// Device/Application/Equipment/FB_VacuumGripper
(*
    FB_VacuumGripper
    Purpose : Suction gripper: valve control with grip and loss supervision.
    Inputs  : xCmdVacuum, xVacuumOk (vacuum switch), tGripTimeout, itfAlarms
    Outputs : xValveOn, xHolding (vacuum on and OK)
    Errors  : VacuumNoGrip - commanded but not OK within tGripTimeout
              VacuumLost - was holding and lost vacuum while still commanded
*)
FUNCTION_BLOCK FB_VacuumGripper IMPLEMENTS I_Equipment
VAR_INPUT
    xCmdVacuum : BOOL;
    xVacuumOk : BOOL;
    tGripTimeout : TIME := T#500MS;
    itfAlarms : I_AlarmSink;
END_VAR
VAR_OUTPUT
    xValveOn : BOOL;
    xHolding : BOOL;
END_VAR
VAR
    tonGrip : TON;
    xWasHolding : BOOL;
    eError : E_AlarmId;
END_VAR

xValveOn := xCmdVacuum;
xHolding := xCmdVacuum AND xVacuumOk;

tonGrip(IN := xCmdVacuum AND NOT xVacuumOk AND NOT xWasHolding, PT := tGripTimeout);
IF tonGrip.Q AND eError = E_AlarmId.None THEN
    eError := E_AlarmId.VacuumNoGrip;
END_IF
IF xWasHolding AND xCmdVacuum AND NOT xVacuumOk AND eError = E_AlarmId.None THEN
    eError := E_AlarmId.VacuumLost;
END_IF

IF xHolding THEN
    xWasHolding := TRUE;
ELSIF NOT xCmdVacuum THEN
    xWasHolding := FALSE;
END_IF

IF eError <> E_AlarmId.None AND itfAlarms <> 0 THEN
    itfAlarms.Raise(eError);
END_IF

METHOD Reset : BOOL
IF itfAlarms <> 0 AND eError <> E_AlarmId.None THEN
    itfAlarms.Clear(eError);
END_IF
eError := E_AlarmId.None;
xWasHolding := FALSE;
Reset := TRUE;
END_METHOD

PROPERTY HasError : BOOL
GET
HasError := eError <> E_AlarmId.None;
END_GET
END_PROPERTY

PROPERTY ErrorId : E_AlarmId
GET
ErrorId := eError;
END_GET
END_PROPERTY

END_FUNCTION_BLOCK

// Device/Application/Equipment/FB_Bin
(*
    FB_Bin
    Purpose : Output bin: counts placed parts and reports the full sensor.
    Inputs  : eBin - which bin; xFullSensor; xPlaced - rising edge = one part placed
    Outputs : uiCount, xFull
    Methods : Empty() - operator emptied the bin
*)
FUNCTION_BLOCK FB_Bin
VAR_INPUT
    eBin : E_Bin;
    xFullSensor : BOOL;
    xPlaced : BOOL;
END_VAR
VAR_OUTPUT
    uiCount : UINT;
    xFull : BOOL;
END_VAR
VAR
    rtPlaced : R_TRIG;
END_VAR

rtPlaced(CLK := xPlaced);
IF rtPlaced.Q THEN
    uiCount := uiCount + 1;
END_IF
xFull := xFullSensor;

METHOD Empty
uiCount := 0;
END_METHOD

END_FUNCTION_BLOCK

// Device/Application/Equipment/FB_PhotoEye
(*
    FB_PhotoEye
    Purpose : Debounced photo-eye with a rising-edge pulse.
    Inputs  : xRaw - sensor signal (TRUE = beam blocked); tDebounce - on/off filter time
    Outputs : xBlocked - debounced state; xRising - TRUE for one cycle when it becomes blocked
*)
FUNCTION_BLOCK FB_PhotoEye
VAR_INPUT
    xRaw : BOOL;
    tDebounce : TIME := T#10MS;
END_VAR
VAR_OUTPUT
    xBlocked : BOOL;
    xRising : BOOL;
END_VAR
VAR
    tonOn : TON;
    tonOff : TON;
END_VAR

tonOn(IN := xRaw, PT := tDebounce);
tonOff(IN := NOT xRaw, PT := tDebounce);
xRising := FALSE;
IF tonOn.Q AND NOT xBlocked THEN
    xBlocked := TRUE;
    xRising := TRUE;
ELSIF tonOff.Q THEN
    xBlocked := FALSE;
END_IF

END_FUNCTION_BLOCK

// Device/Application/Comm/FB_BridgeWatchdog
(*
    FB_BridgeWatchdog
    Purpose : The Python bridge toggles xHeartbeat every cycle; if it stops toggling for tTimeout
              while enabled, the connection to the digital twin is considered lost.
    Outputs : xLost
    Alarms  : BridgeLost (Critical -> the cell aborts)
*)
FUNCTION_BLOCK FB_BridgeWatchdog
VAR_INPUT
    xHeartbeat : BOOL;
    xEnable : BOOL;
    tTimeout : TIME := T#500MS;
    itfAlarms : I_AlarmSink;
END_VAR
VAR_OUTPUT
    xLost : BOOL;
END_VAR
VAR
    xLastHeartbeat : BOOL;
    tonLost : TON;
END_VAR

tonLost(IN := xEnable AND xHeartbeat = xLastHeartbeat, PT := tTimeout);
xLastHeartbeat := xHeartbeat;
xLost := tonLost.Q;
IF itfAlarms <> 0 THEN
    IF xLost THEN
        itfAlarms.Raise(E_AlarmId.BridgeLost);
    ELSE
        itfAlarms.Clear(E_AlarmId.BridgeLost);
    END_IF
END_IF

END_FUNCTION_BLOCK

// Device/Application/Hmi/FB_HmiPanel
(*
    FB_HmiPanel
    Purpose : Turns the operator panel (GVL_HmiPanel: buttons, mode selector) into the cell's
              commands (GVL_Hmi). A button acts on its rising edge and is cleared, so a held or
              stuck button cannot repeat a command; the PackML state machine rejects commands
              that are not allowed in the current state.
    Inputs  : GVL_HmiPanel (written by the visualization), GVL_Bridge.eState
    Outputs : GVL_Hmi.eCommand / eModeRequest / xAlarmAck
    Modes   : iModeSelect 1 Production, 2 Maintenance, 3 Manual; other values are ignored. An
              operator change is requested only where PackML accepts a mode change (Stopped,
              Idle, Aborted), so no request waits to take effect after a later abort. The
              selector then shows GVL_Hmi.eModeRequest, whoever wrote it (panel or OPC UA).
*)
FUNCTION_BLOCK FB_HmiPanel
VAR
    rtStart : R_TRIG;
    rtStop : R_TRIG;
    rtReset : R_TRIG;
    rtClear : R_TRIG;
    rtAbort : R_TRIG;
    rtSuspend : R_TRIG;
    rtUnsuspend : R_TRIG;
    rtAck : R_TRIG;
    iLastMode : INT := 1;  // the selector value the panel showed last cycle
    xModeChangeAllowed : BOOL;
END_VAR

rtStart(CLK := GVL_HmiPanel.xStart);
rtStop(CLK := GVL_HmiPanel.xStop);
rtReset(CLK := GVL_HmiPanel.xReset);
rtClear(CLK := GVL_HmiPanel.xClear);
rtAbort(CLK := GVL_HmiPanel.xAbort);
rtSuspend(CLK := GVL_HmiPanel.xSuspend);
rtUnsuspend(CLK := GVL_HmiPanel.xUnsuspend);
rtAck(CLK := GVL_HmiPanel.xAckAll);

// Abort and Stop first: a safety-relevant command wins over a start in the same cycle.
IF rtAbort.Q THEN
    GVL_Hmi.eCommand := E_PackMLCommand.Abort;
ELSIF rtStop.Q THEN
    GVL_Hmi.eCommand := E_PackMLCommand.Stop;
ELSIF rtClear.Q THEN
    GVL_Hmi.eCommand := E_PackMLCommand.Clear;
ELSIF rtReset.Q THEN
    GVL_Hmi.eCommand := E_PackMLCommand.Reset;
ELSIF rtSuspend.Q THEN
    GVL_Hmi.eCommand := E_PackMLCommand.Suspend;
ELSIF rtUnsuspend.Q THEN
    GVL_Hmi.eCommand := E_PackMLCommand.Unsuspend;
ELSIF rtStart.Q THEN
    GVL_Hmi.eCommand := E_PackMLCommand.Start;
END_IF
IF rtAck.Q THEN
    GVL_Hmi.xAlarmAck := TRUE;
END_IF

// mode selector: an operator change, only where PackML accepts it
IF GVL_HmiPanel.iModeSelect <> iLastMode THEN
    xModeChangeAllowed := GVL_Bridge.eState = E_PackMLState.Stopped
                          OR GVL_Bridge.eState = E_PackMLState.Idle
                          OR GVL_Bridge.eState = E_PackMLState.Aborted;
    IF xModeChangeAllowed THEN
        CASE GVL_HmiPanel.iModeSelect OF
            1: GVL_Hmi.eModeRequest := E_PackMLMode.Production;
            2: GVL_Hmi.eModeRequest := E_PackMLMode.Maintenance;
            3: GVL_Hmi.eModeRequest := E_PackMLMode.Manual;
        END_CASE   // other values: ignored
    END_IF
END_IF
// the selector shows the request (refused or invalid choices fall back, OPC UA requests show)
CASE GVL_Hmi.eModeRequest OF
    E_PackMLMode.Production: iLastMode := 1;
    E_PackMLMode.Maintenance: iLastMode := 2;
    E_PackMLMode.Manual: iLastMode := 3;
END_CASE
GVL_HmiPanel.iModeSelect := iLastMode;

GVL_HmiPanel.xStart := FALSE;
GVL_HmiPanel.xStop := FALSE;
GVL_HmiPanel.xReset := FALSE;
GVL_HmiPanel.xClear := FALSE;
GVL_HmiPanel.xAbort := FALSE;
GVL_HmiPanel.xSuspend := FALSE;
GVL_HmiPanel.xUnsuspend := FALSE;
GVL_HmiPanel.xAckAll := FALSE;

END_FUNCTION_BLOCK

// Device/Application/Hmi/FB_HmiView
(*
    FB_HmiView
    Purpose : Prepares the display data of the visualization (GVL_HmiView): state and mode texts,
              state groups for the machine bar, alarm rows (active or unacknowledged, and the
              condition itself), newest alarm text, equipment signals and the placed counter.
    In/Out  : Cell - the sorting cell (read only)
    Outputs : GVL_HmiView
*)
FUNCTION_BLOCK FB_HmiView
VAR_IN_OUT
    Cell : FB_SortingCell;
END_VAR
VAR
    i : INT;
    stAlarm : ST_Alarm;
END_VAR
VAR CONSTANT
    BELT_RUNNING_MM_S : LREAL := 1.0;  // the belt counts as running above this speed
    // HMI row i shows alarm ALARM_ROWS[i] (E_AlarmId is strict: no integer arithmetic on it)
    ALARM_ROWS : ARRAY[1..16] OF E_AlarmId := [
        E_AlarmId.EStop, E_AlarmId.DoorOpen, E_AlarmId.BridgeLost, E_AlarmId.AxisGroupError,
        E_AlarmId.ConveyorError, E_AlarmId.FollowingErrorWarn, E_AlarmId.FollowingErrorFault,
        E_AlarmId.FeedbackStale, E_AlarmId.VacuumNoGrip, E_AlarmId.VacuumLost,
        E_AlarmId.PartMissed, E_AlarmId.BinFull, E_AlarmId.VisionMissing,
        E_AlarmId.DecisionFallback, E_AlarmId.LowConfidence, E_AlarmId.QueueOverflow];
END_VAR

CASE Cell.eState OF
    E_PackMLState.Clearing: GVL_HmiView.sState := 'Clearing';
    E_PackMLState.Stopped: GVL_HmiView.sState := 'Stopped';
    E_PackMLState.Starting: GVL_HmiView.sState := 'Starting';
    E_PackMLState.Idle: GVL_HmiView.sState := 'Idle';
    E_PackMLState.Suspended: GVL_HmiView.sState := 'Suspended';
    E_PackMLState.Execute: GVL_HmiView.sState := 'Execute';
    E_PackMLState.Stopping: GVL_HmiView.sState := 'Stopping';
    E_PackMLState.Aborting: GVL_HmiView.sState := 'Aborting';
    E_PackMLState.Aborted: GVL_HmiView.sState := 'Aborted';
    E_PackMLState.Holding: GVL_HmiView.sState := 'Holding';
    E_PackMLState.Held: GVL_HmiView.sState := 'Held';
    E_PackMLState.Unholding: GVL_HmiView.sState := 'Unholding';
    E_PackMLState.Suspending: GVL_HmiView.sState := 'Suspending';
    E_PackMLState.Unsuspending: GVL_HmiView.sState := 'Unsuspending';
    E_PackMLState.Resetting: GVL_HmiView.sState := 'Resetting';
    E_PackMLState.Completing: GVL_HmiView.sState := 'Completing';
    E_PackMLState.Complete: GVL_HmiView.sState := 'Complete';
ELSE
    GVL_HmiView.sState := 'Undefined';
END_CASE
CASE Cell.eMode OF
    E_PackMLMode.Production: GVL_HmiView.sMode := 'Production';
    E_PackMLMode.Maintenance: GVL_HmiView.sMode := 'Maintenance';
    E_PackMLMode.Manual: GVL_HmiView.sMode := 'Manual';
END_CASE
CASE Cell.ePickStep OF
    E_PickStep.Idle: GVL_HmiView.sPickStep := 'Idle';
    E_PickStep.MoveHome: GVL_HmiView.sPickStep := 'Moving home';
    E_PickStep.MoveReady: GVL_HmiView.sPickStep := 'Moving to ready';
    E_PickStep.WaitPart: GVL_HmiView.sPickStep := 'Waiting for a part';
    E_PickStep.StartTracking: GVL_HmiView.sPickStep := 'Tracking the belt';
    E_PickStep.Approach: GVL_HmiView.sPickStep := 'Approaching';
    E_PickStep.Descend: GVL_HmiView.sPickStep := 'Descending';
    E_PickStep.Grip: GVL_HmiView.sPickStep := 'Gripping';
    E_PickStep.Lift: GVL_HmiView.sPickStep := 'Lifting';
    E_PickStep.MoveToBin: GVL_HmiView.sPickStep := 'Moving to bin';
    E_PickStep.Release: GVL_HmiView.sPickStep := 'Releasing';
    E_PickStep.Retract: GVL_HmiView.sPickStep := 'Retracting';
    E_PickStep.Aborting: GVL_HmiView.sPickStep := 'Stopping';
    E_PickStep.Aborted: GVL_HmiView.sPickStep := 'Stopped (abort)';
    E_PickStep.Error: GVL_HmiView.sPickStep := 'Error';
    E_PickStep.RecoverLift: GVL_HmiView.sPickStep := 'Recovering';
END_CASE

GVL_HmiView.xExecute := Cell.eState = E_PackMLState.Execute;
GVL_HmiView.xStopped := Cell.eState = E_PackMLState.Stopped;
GVL_HmiView.xIdle := Cell.eState = E_PackMLState.Idle;
GVL_HmiView.xAborted := Cell.eState = E_PackMLState.Aborted OR Cell.eState = E_PackMLState.Aborting;
GVL_HmiView.xHeld := Cell.eState = E_PackMLState.Held OR Cell.eState = E_PackMLState.Suspended
                     OR Cell.eState = E_PackMLState.Holding OR Cell.eState = E_PackMLState.Suspending;
GVL_HmiView.xActing := Cell.eState = E_PackMLState.Resetting OR Cell.eState = E_PackMLState.Starting
                       OR Cell.eState = E_PackMLState.Stopping OR Cell.eState = E_PackMLState.Clearing
                       OR Cell.eState = E_PackMLState.Unholding OR Cell.eState = E_PackMLState.Unsuspending;
GVL_HmiView.xManual := Cell.eMode = E_PackMLMode.Manual;
GVL_HmiView.xJogPermitted := GVL_HmiView.xManual AND GVL_HmiView.xExecute;

GVL_HmiView.xAnyAlarm := FALSE;
FOR i := 1 TO 16 DO
    stAlarm := Cell.AlarmState(ALARM_ROWS[i]);
    GVL_HmiView.axAlarmActive[i] := stAlarm.xActive;
    GVL_HmiView.axAlarm[i] := stAlarm.xActive OR NOT stAlarm.xAcked;
    GVL_HmiView.xAnyAlarm := GVL_HmiView.xAnyAlarm OR GVL_HmiView.axAlarm[i];
END_FOR
GVL_HmiView.sNewestAlarm := GVL_AlarmDefs.aDefs[Cell.eNewestAlarm].sText;
GVL_HmiView.uiPlaced := Cell.PlacedCount();
GVL_HmiView.xBeltRunning := ABS(Cell.lrBeltVel) > BELT_RUNNING_MM_S;
GVL_HmiView.xRobotMoving := Cell.RobotMoving();
GVL_HmiView.xAnyBinFull := Cell.AnyBinFull();

END_FUNCTION_BLOCK

// Device/Application/Tests/PRG_Tests
(*
    PRG_Tests
    Purpose : Calls every simulation test harness (TEST programs in this folder).
    Task    : TestTask, cyclic 10 ms
*)
PROGRAM PRG_Tests
VAR
END_VAR

PRG_TestMotionSmoke();
PRG_TestTypes();
PRG_TestPackML();
PRG_TestAlarms();
PRG_TestEquipment();
PRG_TestMotion();
PRG_TestJointMonitor();
PRG_TestTracking();
PRG_TestPick();
PRG_TestCell();

END_PROGRAM

// Device/Application/Tests/PRG_TestMotionSmoke
(*
    PRG_TestMotionSmoke
    Purpose : Simulation test harness - powers the robot axis group and makes one PTP move.
    Task    : TestTask (via PRG_Tests)
    Spec    : tests/plc/motion_smoke.json
*)
PROGRAM PRG_TestMotionSmoke
VAR
    fbPower : SMC_GroupPower;
    fbEnable : MC_GroupEnable;
    fbMove : MC_MoveDirectAbsolute := (CoordSystem := SMC_COORD_SYSTEM.ACS, VelFactor := 0.5);
    fbReadPos : MC_GroupReadActualPosition := (Enable := TRUE, CoordSystem := SMC_COORD_SYSTEM.ACS);
    xGo : BOOL;
    lrJ1 : LREAL;
    lrJ2 : LREAL;
    xMoveDone : BOOL;
    xMoveError : BOOL;
END_VAR

// Only commands the robot while the test runs, so other harnesses can use it.
IF xGo THEN
    fbPower(AxisGroup := AxisGroup_Robot, Enable := TRUE, bRegulatorOn := TRUE, bDriveStart := TRUE);
    fbEnable(AxisGroup := AxisGroup_Robot, Execute := fbPower.Status);
    fbMove.Position.a.a0 := 30;
    fbMove.Position.a.a1 := -20;
    fbMove.Position.a.a2 := 40;
    fbMove.Position.a.a3 := 0;
    fbMove.Position.a.a4 := 45;
    fbMove.Position.a.a5 := 0;
    fbMove(AxisGroup := AxisGroup_Robot, Execute := fbEnable.Done);
    fbReadPos(AxisGroup := AxisGroup_Robot);
    lrJ1 := fbReadPos.Position.a.a0;
    lrJ2 := fbReadPos.Position.a.a1;
    xMoveDone := fbMove.Done;
    xMoveError := fbMove.Error;
END_IF

END_PROGRAM

// Device/Application/Tests/PRG_TestTypes
(*
    PRG_TestTypes
    Purpose : Simulation test harness - exposes configuration values for tests/plc/types.json.
*)
PROGRAM PRG_TestTypes
VAR
    eClassBin0 : E_Bin;
    eFaultClass : E_AlarmClass;
    eWarnClass : E_AlarmClass;
    xLoopback : BOOL;
END_VAR

eClassBin0 := GVL_Params.aClassToBin[0];
eFaultClass := GVL_AlarmDefs.aDefs[E_AlarmId.EStop].eClass;
eWarnClass := GVL_AlarmDefs.aDefs[E_AlarmId.PartMissed].eClass;
xLoopback := GVL_Config.xFeedbackLoopback;

END_PROGRAM

// Device/Application/Tests/PRG_TestPackML
(*
    PRG_TestPackML
    Purpose : Simulation test harness for FB_PackMLStateMachine (tests/plc/packml.json).
    Inputs  : xReinit - TRUE re-initialises the state machine, then resets itself.
*)
PROGRAM PRG_TestPackML
VAR
    fbSm : FB_PackMLStateMachine;
    fbSmInitial : FB_PackMLStateMachine;
    xReinit : BOOL;
END_VAR

IF xReinit THEN
    xReinit := FALSE;
    fbSm := fbSmInitial;
END_IF
fbSm();

END_PROGRAM

// Device/Application/Tests/PRG_TestAlarms
(*
    PRG_TestAlarms
    Purpose : Simulation test harness for FB_AlarmHandler (tests/plc/alarms.json).
    Inputs  : eId + xRaise / xRaiseEvent / xClear pulses, xAck, xReinit (each pulse resets itself).
*)
PROGRAM PRG_TestAlarms
VAR
    fbAlarms : FB_AlarmHandler;
    fbAlarmsInitial : FB_AlarmHandler;
    eId : E_AlarmId;
    xRaise : BOOL;
    xRaiseEvent : BOOL;
    xClear : BOOL;
    xAck : BOOL;
    xReinit : BOOL;
END_VAR

IF xReinit THEN
    xReinit := FALSE;
    fbAlarms := fbAlarmsInitial;
END_IF
IF xRaise THEN
    xRaise := FALSE;
    fbAlarms.Raise(eId);
END_IF
IF xRaiseEvent THEN
    xRaiseEvent := FALSE;
    fbAlarms.RaiseEvent(eId);
END_IF
IF xClear THEN
    xClear := FALSE;
    fbAlarms.Clear(eId);
END_IF
IF xAck THEN
    xAck := FALSE;
    fbAlarms.AcknowledgeAll();
END_IF
fbAlarms();

END_PROGRAM

// Device/Application/Tests/PRG_TestEquipment
(*
    PRG_TestEquipment
    Purpose : Simulation test harness for the simple equipment FBs (tests/plc/equipment.json).
    Pulses  : write udiPulseMs and set xStartPulse - the harness drives fbPe.xRaw for exactly
              that long in PLC time (tool writes are too slow to time a short pulse).
*)
PROGRAM PRG_TestEquipment
VAR
    fbAlarms : FB_AlarmHandler;
    fbPe : FB_PhotoEye := (tDebounce := T#300MS);
    fbVac : FB_VacuumGripper;
    fbBin : FB_Bin := (eBin := E_Bin.TypeA);
    fbSafety : FB_SafetyMonitor;
    fbAlarmsInitial : FB_AlarmHandler;
    fbPeInitial : FB_PhotoEye := (tDebounce := T#300MS);
    fbVacInitial : FB_VacuumGripper;
    fbBinInitial : FB_Bin := (eBin := E_Bin.TypeA);
    fbSafetyInitial : FB_SafetyMonitor;
    xReinit : BOOL;
    uiPeRises : UINT;
    eVacError : E_AlarmId;
    udiPulseMs : UDINT;
    xStartPulse : BOOL;
    xPulseActive : BOOL;
    tonPulse : TON;
END_VAR

IF xReinit THEN
    xReinit := FALSE;
    fbAlarms := fbAlarmsInitial;
    fbPe := fbPeInitial;
    fbVac := fbVacInitial;
    fbBin := fbBinInitial;
    fbSafety := fbSafetyInitial;
    uiPeRises := 0;
    xPulseActive := FALSE;
END_IF
fbVac.itfAlarms := fbAlarms;
fbSafety.itfAlarms := fbAlarms;

IF xStartPulse THEN
    xStartPulse := FALSE;
    xPulseActive := TRUE;
END_IF
tonPulse(IN := xPulseActive, PT := TO_TIME(udiPulseMs));
IF tonPulse.Q THEN
    xPulseActive := FALSE;
END_IF
fbPe.xRaw := xPulseActive;

fbPe();
IF fbPe.xRising THEN
    uiPeRises := uiPeRises + 1;
END_IF
fbVac();
eVacError := fbVac.ErrorId;
fbBin();
fbSafety();
fbAlarms();

END_PROGRAM

// Device/Application/Tests/PRG_TestMotion
(*
    PRG_TestMotion
    Purpose : Simulation test harness for FB_Robot and FB_Conveyor (tests/plc/motion.json).
    Inputs  : xActive - only then are the FBs called; xGo - start eCmd with the target chosen by
              iTargetSel (1 = home, 2 = current TCP - 50 mm in Z, 3 = home with J1 = 60 deg,
              4 = stProbe as written by the test)
    Outputs : xLastDone / xLastError of the last command, udiMoveMsLast / udiMoveMsPrev,
              xSlower (last move took > 1.5 x the previous one), lrZDelta
    Note    : SoftMotion FB instances are never re-initialised by assignment (corrupts them).
*)
PROGRAM PRG_TestMotion
VAR
    fbRobot : FB_Robot;
    fbConv : FB_Conveyor;
    fbAlarms : FB_AlarmHandler;
    xActive : BOOL;
    iTargetSel : INT;
    eCmd : E_RobotCmd;
    xGo : BOOL;
    iGoStep : INT;
    xLastDone : BOOL;
    xLastError : BOOL;
    tStart : TIME;
    udiMoveMsLast : UDINT;
    udiMoveMsPrev : UDINT;
    xSlower : BOOL;
    lrZStart : LREAL;
    lrZDelta : LREAL;
    stTarget : SMC_POS_REF;
    stProbe : SMC_POS_REF;
END_VAR

IF NOT xActive THEN
    RETURN;
END_IF
fbRobot.itfAlarms := fbAlarms;
fbConv.itfAlarms := fbAlarms;

IF xGo THEN
    xGo := FALSE;
    CASE iTargetSel OF
        1: stTarget := GVL_CellGeometry.HOME_ACS;
        2: stTarget := fbRobot.stActMcs;
           lrZStart := fbRobot.stActMcs.c.Z;
           stTarget.c.Z := lrZStart - 50;
        3: stTarget := GVL_CellGeometry.HOME_ACS;
           stTarget.a.a0 := 60;
        4: stTarget := stProbe;
    END_CASE
    fbRobot.stTarget := stTarget;
    fbRobot.eCmd := eCmd;
    fbRobot.xExecute := FALSE;     // a fresh rising edge, even if a command is running
    iGoStep := 1;
    xLastDone := FALSE;
    xLastError := FALSE;
ELSIF iGoStep = 1 THEN
    fbRobot.xExecute := TRUE;
    tStart := TIME();
    iGoStep := 2;
ELSIF iGoStep = 2 AND (fbRobot.xDone OR fbRobot.xError) THEN
    xLastDone := fbRobot.xDone;
    xLastError := fbRobot.xError;
    udiMoveMsPrev := udiMoveMsLast;
    udiMoveMsLast := TIME_TO_UDINT(TIME() - tStart);
    xSlower := udiMoveMsLast * 2 > udiMoveMsPrev * 3;
    fbRobot.xExecute := FALSE;
    iGoStep := 0;
END_IF

fbRobot(AxisGroup := AxisGroup_Robot);
fbConv(Axis := Axis_Conveyor);
fbAlarms();
IF iTargetSel = 2 THEN
    lrZDelta := fbRobot.stActMcs.c.Z - lrZStart;
END_IF

END_PROGRAM

// Device/Application/Tests/PRG_TestJointMonitor
(*
    PRG_TestJointMonitor
    Purpose : Simulation test harness for FB_JointMonitor (tests/plc/joint_monitor.json).
    Inputs  : xReinit; xAutoSeq - increment the feedback and setpoint sequences every cycle
              xRamp - J1 setpoint ramps by RAMP_STEP per cycle; iLag - feedback is the setpoint of
              iLag cycles earlier (and says so in udiFeedbackForSeq); xFreeze - feedback stands still;
              iTornSamples - that many cycles claim a sample iTornAge older (a torn OPC UA write,
              or a bridge hiccup when iTornAge exceeds the history)
    Outputs : lrRampSpeed - measured J1 setpoint speed [deg/s]
*)
PROGRAM PRG_TestJointMonitor
VAR
    fbMon : FB_JointMonitor;
    fbAlarms : FB_AlarmHandler;
    fbMonInitial : FB_JointMonitor;
    fbAlarmsInitial : FB_AlarmHandler;
    xReinit : BOOL;
    xAutoSeq : BOOL;
    xRamp : BOOL;
    xFreeze : BOOL;
    iLag : INT;
    udiSpSeq : UDINT;
    aSpHist : ARRAY[0..127] OF LREAL;
    xRampOld : BOOL;
    tRampStart : TIME;
    lrRampStart : LREAL;
    lrRampSpeed : LREAL;
    iTornSamples : INT;             // next cycles: feedback says it answers an older sample
    iTornAge : INT := 25;           // [samples]
END_VAR
VAR CONSTANT
    RAMP_STEP : LREAL := 1.0;       // [deg per cycle]
END_VAR

IF xReinit THEN
    xReinit := FALSE;
    xAutoSeq := FALSE;
    xRamp := FALSE;
    xFreeze := FALSE;
    iLag := 0;
    iTornSamples := 0;
    udiSpSeq := 0;
    fbMon := fbMonInitial;
    fbAlarms := fbAlarmsInitial;
END_IF
IF xAutoSeq THEN
    fbMon.udiFeedbackSeq := fbMon.udiFeedbackSeq + 1;
    udiSpSeq := udiSpSeq + 1;
END_IF
IF xRamp THEN
    IF NOT xRampOld THEN
        tRampStart := TIME();
        lrRampStart := fbMon.aSetpoint[1];
    END_IF
    fbMon.aSetpoint[1] := fbMon.aSetpoint[1] + RAMP_STEP;
    IF TIME() > tRampStart THEN
        lrRampSpeed := (fbMon.aSetpoint[1] - lrRampStart) * 1000.0 / TIME_TO_LREAL(TIME() - tRampStart);
    END_IF
END_IF
xRampOld := xRamp;
aSpHist[udiSpSeq MOD 128] := fbMon.aSetpoint[1];
fbMon.udiSetpointSeq := udiSpSeq;
IF udiSpSeq >= INT_TO_UDINT(iLag) THEN
    fbMon.udiFeedbackForSeq := udiSpSeq - INT_TO_UDINT(iLag);
    IF NOT xFreeze THEN
        fbMon.aFeedback[1] := aSpHist[fbMon.udiFeedbackForSeq MOD 128];
    END_IF
    IF iTornSamples > 0 AND fbMon.udiFeedbackForSeq >= INT_TO_UDINT(iTornAge) THEN
        fbMon.udiFeedbackForSeq := fbMon.udiFeedbackForSeq - INT_TO_UDINT(iTornAge);
        iTornSamples := iTornSamples - 1;
    END_IF
END_IF
fbMon.itfAlarms := fbAlarms;
fbMon();
fbAlarms();

END_PROGRAM

// Device/Application/Tests/PRG_TestTracking
(*
    PRG_TestTracking
    Purpose : Simulation test harness for FB_PartTracker and F_SelectBin (tests/plc/tracking.json).
    Inputs  : lrBeltPos; xTriggerPE1 (one capture); uiFillCount (that many captures, one per cycle);
              stVisIn + xSendVision / xResendVision (same sequence number again);
              stDecIn + xSendDecision; udiQueryId - part to show in stRec; xAck; xClear;
              xNoDecisionLayer (no AI decision service)
    Outputs : uiCount, uiNext (next pickable index), stRec, xQueryFound
*)
PROGRAM PRG_TestTracking
VAR
    fbTracker : FB_PartTracker;
    fbAlarms : FB_AlarmHandler;
    fbTrackerInitial : FB_PartTracker;
    fbAlarmsInitial : FB_AlarmHandler;
    xReinit : BOOL;
    lrBeltPos : LREAL;
    xTriggerPE1 : BOOL;
    uiFillCount : UINT;
    stVisIn : ST_VisionMsg;
    stDecIn : ST_DecisionMsg;
    xSendVision : BOOL;
    xResendVision : BOOL;
    xSendDecision : BOOL;
    xAck : BOOL;
    xClear : BOOL;
    udiVisionSeq : UDINT;
    udiDecisionSeq : UDINT;
    udiQueryId : UDINT;
    uiQueryIdx : UINT;
    xQueryFound : BOOL;
    stRec : ST_PartRecord;
    uiCount : UINT;
    uiNext : UINT;
    xPE1Rising : BOOL;
    xNoDecisionLayer : BOOL;
END_VAR

IF xReinit THEN
    xReinit := FALSE;
    fbTracker := fbTrackerInitial;
    fbAlarms := fbAlarmsInitial;
    udiVisionSeq := 0;
    udiDecisionSeq := 0;
    uiFillCount := 0;
END_IF

xPE1Rising := xTriggerPE1 OR uiFillCount > 0;
xTriggerPE1 := FALSE;
IF uiFillCount > 0 THEN
    uiFillCount := uiFillCount - 1;
END_IF

IF xSendVision THEN
    xSendVision := FALSE;
    udiVisionSeq := udiVisionSeq + 1;
END_IF
IF xResendVision THEN
    xResendVision := FALSE;      // same sequence number: must be ignored
END_IF
stVisIn.udiSeq := udiVisionSeq;
IF xSendDecision THEN
    xSendDecision := FALSE;
    udiDecisionSeq := udiDecisionSeq + 1;
END_IF
stDecIn.udiSeq := udiDecisionSeq;
IF xAck THEN
    xAck := FALSE;
    fbAlarms.AcknowledgeAll();
END_IF
IF xClear THEN
    xClear := FALSE;
    fbTracker.Clear();
END_IF

fbTracker.itfAlarms := fbAlarms;
fbTracker(lrBeltPos := lrBeltPos, xPE1Rising := xPE1Rising, stVision := stVisIn, stDecision := stDecIn,
          xDecisionActive := NOT xNoDecisionLayer);
fbAlarms();

uiCount := fbTracker.Count;
uiNext := fbTracker.NextPickable(GVL_CellGeometry.PE2_X, GVL_CellGeometry.PICK_WINDOW_END_X);
uiQueryIdx := fbTracker.FindPart(udiQueryId);
xQueryFound := uiQueryIdx > 0;
IF xQueryFound THEN
    stRec := fbTracker.GetRecord(uiQueryIdx);
END_IF

END_PROGRAM

// Device/Application/Tests/PRG_TestPick
(*
    PRG_TestPick
    Purpose : Simulation test harness for FB_PickSequence (tests/plc/pick.json). Owns the robot,
              conveyor, gripper, tracker and alarms like the cell does, and simulates the vacuum
              switch (OK 100 ms after the valve opens).
    Inputs  : xActive, xBeltRun, xInject (+ usiInjClass, eInjQuality, lrInjX: one part with
              vision and decision; xInjInvalid: the vision message says "not seen"),
              xDropOnTransfer (vacuum lost during MoveToBin),
              xAbortOnLift (abort when the sequence reaches Lift), xResetSeq
    Outputs : xSawRecoverLift (latched: the recovery after an abort lifted first),
              lrGripZ (TCP height when the last grip started) [mm]
    Note    : SoftMotion FB instances are never re-initialised by assignment.
*)
PROGRAM PRG_TestPick
VAR
    fbRobot : FB_Robot;
    fbConv : FB_Conveyor;
    fbVac : FB_VacuumGripper;
    fbTracker : FB_PartTracker;
    fbAlarms : FB_AlarmHandler;
    fbSeq : FB_PickSequence;
    xActive : BOOL;
    xBeltRun : BOOL;
    xInject : BOOL;
    xInjInvalid : BOOL;
    usiInjClass : USINT;
    eInjQuality : E_Quality := E_Quality.Ok;
    lrInjX : LREAL := 1000;
    iInject : INT;
    xPE1 : BOOL;
    stVis : ST_VisionMsg;
    stDec : ST_DecisionMsg;
    xDropOnTransfer : BOOL;
    xAbortOnLift : BOOL;
    xResetSeq : BOOL;
    xVacLost : BOOL;
    tonVac : TON;
    xSawRecoverLift : BOOL;
    lrGripZ : LREAL;
    eLastStep : E_PickStep;
END_VAR

IF NOT xActive THEN
    RETURN;
END_IF
fbRobot.itfAlarms := fbAlarms;
fbConv.itfAlarms := fbAlarms;
fbVac.itfAlarms := fbAlarms;
fbTracker.itfAlarms := fbAlarms;
fbConv.xEnable := TRUE;
fbConv.lrVelocity := GVL_Params.lrBeltSpeed;
fbConv.xRun := xBeltRun;
fbRobot.xEnable := TRUE;

// One injected part: capture, then vision, then decision on consecutive cycles.
CASE iInject OF
    0:
        IF xInject THEN
            xInject := FALSE;
            xPE1 := TRUE;
            iInject := 1;
        END_IF
    1:
        xPE1 := FALSE;
        iInject := 2;
    2:
        stVis.udiSeq := stVis.udiSeq + 1;
        stVis.udiPartId := fbTracker.stCapture.udiPartId;
        stVis.xValid := NOT xInjInvalid;
        stVis.usiClass := usiInjClass;
        stVis.rConfidence := 0.9;
        stVis.lrX := lrInjX;
        stVis.lrY := 0;
        stVis.lrTheta := 0;
        iInject := 3;
    3:
        stDec.udiSeq := stDec.udiSeq + 1;
        stDec.udiPartId := stVis.udiPartId;
        stDec.eQuality := eInjQuality;
        stDec.rQualityProb := 0.95;
        stDec.xIdentReliable := TRUE;
        iInject := 0;
END_CASE

IF xDropOnTransfer AND fbSeq.eStep = E_PickStep.MoveToBin THEN
    xVacLost := TRUE;
END_IF
tonVac(IN := fbVac.xValveOn AND NOT xVacLost, PT := T#100MS);
fbVac.xVacuumOk := tonVac.Q;
IF xAbortOnLift AND fbSeq.eStep = E_PickStep.Lift THEN
    fbSeq.xAbort := TRUE;
END_IF
fbSeq.xReset := xResetSeq;
IF xResetSeq THEN
    xResetSeq := FALSE;
    xVacLost := FALSE;
    fbSeq.xAbort := FALSE;
    fbVac.Reset();
    fbAlarms.AcknowledgeAll();
END_IF

fbTracker(lrBeltPos := fbConv.lrPosition, xPE1Rising := xPE1, stVision := stVis, stDecision := stDec);
fbSeq(AxisGroup := AxisGroup_Robot, ConveyorAxis := Axis_Conveyor, Robot := fbRobot, Gripper := fbVac, Tracker := fbTracker);
fbVac();
fbRobot(AxisGroup := AxisGroup_Robot);
fbConv(Axis := Axis_Conveyor);
fbAlarms();
IF fbSeq.eStep = E_PickStep.RecoverLift THEN
    xSawRecoverLift := TRUE;
END_IF
IF fbSeq.eStep = E_PickStep.Grip AND eLastStep <> E_PickStep.Grip THEN
    lrGripZ := fbRobot.stActMcs.c.Z;
END_IF
eLastStep := fbSeq.eStep;

END_PROGRAM

// Device/Application/Tests/PRG_TestCell
(*
    PRG_TestCell
    Purpose : Simulation test harness for the whole cell in PRG_Main (tests/plc/cell.json).
              Simulates the vacuum switch, injects parts (PE1 pulse, then vision and decision
              messages for the captured part id) and can press the E-stop or lose the vacuum
              during a transfer. Can play the twin's bridge (heartbeat, joint feedback answering
              the current setpoint sample, twin active) and stall it. While active it plays an AI
              decision service (GVL_Bridge.xDecisionActive), reset when it is switched off.
    Inputs  : xActive; xInject (+ usiInjClass, eInjQuality); xEStopOnTransfer; xVacLostOnTransfer;
              xMark (J1 reference); xBridgeSim; xBridgeStall (heartbeat stops toggling);
              xBridgeStallOnTransfer
    Outputs : lrJ1Delta - J1 movement since xMark [deg]; lrAbortDelayMs - bridge stall -> Aborted
*)
PROGRAM PRG_TestCell
VAR
    xActive : BOOL;
    xWasActive : BOOL;
    xInject : BOOL;
    usiInjClass : USINT;
    eInjQuality : E_Quality := E_Quality.Ok;
    iInject : INT;
    tonPulse : TON;
    tonVac : TON;
    xEStopOnTransfer : BOOL;
    xVacLostOnTransfer : BOOL;
    xVacLost : BOOL;                    // latched until xVacLostOnTransfer is released
    xMark : BOOL;
    lrJ1Start : LREAL;
    lrJ1Delta : LREAL;
    xBridgeSim : BOOL;
    xBridgeStall : BOOL;
    xBridgeStallOnTransfer : BOOL;      // stall the bridge when the robot carries a part to its bin
    xStallTimed : BOOL;
    tStall : TIME;
    lrAbortDelayMs : LREAL;             // stall -> Aborted [ms]
END_VAR
VAR CONSTANT
    PE1_PULSE : TIME := T#250MS;
END_VAR

IF NOT xActive THEN
    IF xWasActive THEN                   // leave no fake decision service behind
        GVL_Bridge.xDecisionActive := FALSE;
        xWasActive := FALSE;
    END_IF
    RETURN;
END_IF
xWasActive := TRUE;
GVL_Bridge.xDecisionActive := TRUE;  // the harness injects AI decisions (eInjQuality)

IF xVacLostOnTransfer AND PRG_Main.fbCell.ePickStep = E_PickStep.MoveToBin THEN
    xVacLost := TRUE;
ELSIF NOT xVacLostOnTransfer THEN
    xVacLost := FALSE;
END_IF
tonVac(IN := GVL_Bridge.xVacuumOn, PT := T#100MS);
GVL_Bridge.xVacuumOk := tonVac.Q AND NOT xVacLost;

// the twin's bridge: feedback answers the current setpoint sample, heartbeat toggles
IF xBridgeStallOnTransfer AND NOT xBridgeStall AND PRG_Main.fbCell.ePickStep = E_PickStep.MoveToBin THEN
    xBridgeStall := TRUE;
    xStallTimed := FALSE;
    tStall := TIME();
END_IF
IF xBridgeStall AND NOT xStallTimed AND GVL_Bridge.eState = E_PackMLState.Aborted THEN
    xStallTimed := TRUE;
    lrAbortDelayMs := TIME_TO_LREAL(TIME() - tStall);
END_IF
IF xBridgeSim THEN
    GVL_Bridge.xTwinActive := TRUE;
    GVL_Bridge.aJointPosFb := GVL_Bridge.aJointPosSp;
    GVL_Bridge.udiFeedbackForSeq := GVL_Bridge.udiSetpointSeq;
    IF NOT xBridgeStall THEN
        GVL_Bridge.xHeartbeat := NOT GVL_Bridge.xHeartbeat;
        GVL_Bridge.udiFeedbackSeq := GVL_Bridge.udiFeedbackSeq + 1;
    END_IF
END_IF

CASE iInject OF
    0:
        IF xInject THEN
            xInject := FALSE;
            GVL_Bridge.xPE1 := TRUE;
            iInject := 1;
        END_IF
    1:
        tonPulse(IN := TRUE, PT := PE1_PULSE);
        IF tonPulse.Q THEN
            tonPulse(IN := FALSE);
            GVL_Bridge.xPE1 := FALSE;
            iInject := 2;
        END_IF
    2:
        GVL_Bridge.stVision.udiPartId := GVL_Bridge.stCapture.udiPartId;
        GVL_Bridge.stVision.xValid := TRUE;
        GVL_Bridge.stVision.usiClass := usiInjClass;
        GVL_Bridge.stVision.rConfidence := 0.9;
        GVL_Bridge.stVision.lrX := GVL_CellGeometry.PE1_X;
        GVL_Bridge.stVision.lrY := 0;
        GVL_Bridge.stVision.lrTheta := 0;
        GVL_Bridge.stVision.udiSeq := GVL_Bridge.stVision.udiSeq + 1;
        iInject := 3;
    3:
        GVL_Bridge.stDecision.udiPartId := GVL_Bridge.stVision.udiPartId;
        GVL_Bridge.stDecision.eQuality := eInjQuality;
        GVL_Bridge.stDecision.rQualityProb := 0.95;
        GVL_Bridge.stDecision.xIdentReliable := TRUE;
        GVL_Bridge.stDecision.udiSeq := GVL_Bridge.stDecision.udiSeq + 1;
        iInject := 0;
END_CASE

IF xEStopOnTransfer AND PRG_Main.fbCell.ePickStep = E_PickStep.MoveToBin THEN
    GVL_Bridge.xEStopOk := FALSE;
END_IF

IF xMark THEN
    xMark := FALSE;
    lrJ1Start := PRG_Main.fbCell.aActAcs[1];
END_IF
lrJ1Delta := PRG_Main.fbCell.aActAcs[1] - lrJ1Start;

END_PROGRAM

// Device/Application/PRG_Recipe_Cell
PROGRAM PRG_Recipe_Cell
// Set iApply to a recipe's index to write it to the variables; set iSave to store the variables in it.
VAR
    iApply : INT := -1;
    iSave : INT := -1;
    iActive : INT := -1; // the recipe applied last
    sActive : STRING(32);
    p0 : POINTER TO LREAL; // GVL_Params.lrBeltSpeed
    p1 : POINTER TO LREAL; // GVL_Params.lrApproachHeight
    p2 : POINTER TO LREAL; // GVL_Params.lrPickDepth
    p3 : POINTER TO LREAL; // GVL_Params.lrLinVelocity
    p4 : POINTER TO LREAL; // GVL_Params.lrLinAccel
    p5 : POINTER TO LREAL; // GVL_Params.lrLinJerk
    p6 : POINTER TO LREAL; // GVL_Params.lrPtpVelFactor
    p7 : POINTER TO REAL; // GVL_Params.rConfidenceThreshold
    p8 : POINTER TO TIME; // GVL_Params.tDecisionDeadline
    p9 : POINTER TO TIME; // GVL_Params.tVacuumTimeout
    p10 : POINTER TO LREAL; // GVL_Params.lrFollowErrWarn
    p11 : POINTER TO LREAL; // GVL_Params.lrFollowErrFault
    p12 : POINTER TO TIME; // GVL_Params.tFeedbackTimeout
END_VAR

p0 := ADR(GVL_Params.lrBeltSpeed);
p1 := ADR(GVL_Params.lrApproachHeight);
p2 := ADR(GVL_Params.lrPickDepth);
p3 := ADR(GVL_Params.lrLinVelocity);
p4 := ADR(GVL_Params.lrLinAccel);
p5 := ADR(GVL_Params.lrLinJerk);
p6 := ADR(GVL_Params.lrPtpVelFactor);
p7 := ADR(GVL_Params.rConfidenceThreshold);
p8 := ADR(GVL_Params.tDecisionDeadline);
p9 := ADR(GVL_Params.tVacuumTimeout);
p10 := ADR(GVL_Params.lrFollowErrWarn);
p11 := ADR(GVL_Params.lrFollowErrFault);
p12 := ADR(GVL_Params.tFeedbackTimeout);
IF iApply >= 0 AND iApply < 2 THEN
    p0^ := GVL_Recipe_Cell.aRecipes[iApply].lrBeltSpeed;
    p1^ := GVL_Recipe_Cell.aRecipes[iApply].lrApproachHeight;
    p2^ := GVL_Recipe_Cell.aRecipes[iApply].lrPickDepth;
    p3^ := GVL_Recipe_Cell.aRecipes[iApply].lrLinVelocity;
    p4^ := GVL_Recipe_Cell.aRecipes[iApply].lrLinAccel;
    p5^ := GVL_Recipe_Cell.aRecipes[iApply].lrLinJerk;
    p6^ := GVL_Recipe_Cell.aRecipes[iApply].lrPtpVelFactor;
    p7^ := GVL_Recipe_Cell.aRecipes[iApply].rConfidenceThreshold;
    p8^ := GVL_Recipe_Cell.aRecipes[iApply].tDecisionDeadline;
    p9^ := GVL_Recipe_Cell.aRecipes[iApply].tVacuumTimeout;
    p10^ := GVL_Recipe_Cell.aRecipes[iApply].lrFollowErrWarn;
    p11^ := GVL_Recipe_Cell.aRecipes[iApply].lrFollowErrFault;
    p12^ := GVL_Recipe_Cell.aRecipes[iApply].tFeedbackTimeout;
    iActive := iApply;
    sActive := GVL_Recipe_Cell.asNames[iApply];
END_IF
iApply := -1;
IF iSave >= 0 AND iSave < 2 THEN
    GVL_Recipe_Cell.aRecipes[iSave].lrBeltSpeed := p0^;
    GVL_Recipe_Cell.aRecipes[iSave].lrApproachHeight := p1^;
    GVL_Recipe_Cell.aRecipes[iSave].lrPickDepth := p2^;
    GVL_Recipe_Cell.aRecipes[iSave].lrLinVelocity := p3^;
    GVL_Recipe_Cell.aRecipes[iSave].lrLinAccel := p4^;
    GVL_Recipe_Cell.aRecipes[iSave].lrLinJerk := p5^;
    GVL_Recipe_Cell.aRecipes[iSave].lrPtpVelFactor := p6^;
    GVL_Recipe_Cell.aRecipes[iSave].rConfidenceThreshold := p7^;
    GVL_Recipe_Cell.aRecipes[iSave].tDecisionDeadline := p8^;
    GVL_Recipe_Cell.aRecipes[iSave].tVacuumTimeout := p9^;
    GVL_Recipe_Cell.aRecipes[iSave].lrFollowErrWarn := p10^;
    GVL_Recipe_Cell.aRecipes[iSave].lrFollowErrFault := p11^;
    GVL_Recipe_Cell.aRecipes[iSave].tFeedbackTimeout := p12^;
END_IF
iSave := -1;

END_PROGRAM

// Device/Application/PRG_HMI_Alarms
PROGRAM PRG_HMI_Alarms
// Generated by codesys-mcp-toolkit for the HMI screen 'Alarms' (42 variables). Rebuilt on every export.
VAR
    iMachine : INT; // the machine's state: 0 idle, 1.. the states in order
    sV1 : STRING(80); // GVL_HmiView.sState
    sV2 : STRING(80); // GVL_HmiView.sMode
    rV3 : REAL; // GVL_HmiView.sNewestAlarm
END_VAR

IF GVL_HmiView.xAborted THEN iMachine := 1; ELSIF GVL_HmiView.xHeld THEN iMachine := 2; ELSIF GVL_HmiView.xActing THEN iMachine := 3; ELSIF GVL_HmiView.xManual THEN iMachine := 4; ELSIF GVL_HmiView.xExecute THEN iMachine := 5; ELSIF GVL_HmiView.xIdle THEN iMachine := 6; ELSE iMachine := 0; END_IF
sV1 := TO_STRING(GVL_HmiView.sState);
sV2 := TO_STRING(GVL_HmiView.sMode);
rV3 := ANY_TO_REAL(GVL_HmiView.sNewestAlarm);

END_PROGRAM

// Device/Application/PRG_HMI_Robot
PROGRAM PRG_HMI_Robot
// Generated by codesys-mcp-toolkit for the HMI screen 'Robot' (49 variables). Rebuilt on every export.
VAR
    iMachine : INT; // the machine's state: 0 idle, 1.. the states in order
    sV1 : STRING(80); // GVL_HmiView.sState
    sV2 : STRING(80); // GVL_HmiView.sMode
    rV3 : REAL; // GVL_HmiView.uiPlaced
    rV4 : REAL; // GVL_Bridge.aJointPosSp[1]
    iP5 : INT; // GVL_Bridge.aJointPosSp[1]
    rV6 : REAL; // GVL_Bridge.aJointPosSp[2]
    iP7 : INT; // GVL_Bridge.aJointPosSp[2]
    rV8 : REAL; // GVL_Bridge.aJointPosSp[3]
    iP9 : INT; // GVL_Bridge.aJointPosSp[3]
    rV10 : REAL; // GVL_Bridge.aJointPosSp[4]
    iP11 : INT; // GVL_Bridge.aJointPosSp[4]
    rV12 : REAL; // GVL_Bridge.aJointPosSp[5]
    iP13 : INT; // GVL_Bridge.aJointPosSp[5]
    rV14 : REAL; // GVL_Bridge.aJointPosSp[6]
    iP15 : INT; // GVL_Bridge.aJointPosSp[6]
    rV16 : REAL; // GVL_Bridge.aFollowingError[1]
    xB17 : BOOL; // GVL_Bridge.aFollowingError[1] >= 2
    iP18 : INT; // GVL_Bridge.aFollowingError[1]
    xB19 : BOOL; // GVL_Bridge.aFollowingError[1] >= 2
    rV20 : REAL; // GVL_Bridge.aFollowingError[2]
    xB21 : BOOL; // GVL_Bridge.aFollowingError[2] >= 2
    iP22 : INT; // GVL_Bridge.aFollowingError[2]
    xB23 : BOOL; // GVL_Bridge.aFollowingError[2] >= 2
    rV24 : REAL; // GVL_Bridge.aFollowingError[3]
    xB25 : BOOL; // GVL_Bridge.aFollowingError[3] >= 2
    iP26 : INT; // GVL_Bridge.aFollowingError[3]
    xB27 : BOOL; // GVL_Bridge.aFollowingError[3] >= 2
    rV28 : REAL; // GVL_Bridge.aFollowingError[4]
    xB29 : BOOL; // GVL_Bridge.aFollowingError[4] >= 2
    iP30 : INT; // GVL_Bridge.aFollowingError[4]
    xB31 : BOOL; // GVL_Bridge.aFollowingError[4] >= 2
    rV32 : REAL; // GVL_Bridge.aFollowingError[5]
    xB33 : BOOL; // GVL_Bridge.aFollowingError[5] >= 2
    iP34 : INT; // GVL_Bridge.aFollowingError[5]
    xB35 : BOOL; // GVL_Bridge.aFollowingError[5] >= 2
    rV36 : REAL; // GVL_Bridge.aFollowingError[6]
    xB37 : BOOL; // GVL_Bridge.aFollowingError[6] >= 2
    iP38 : INT; // GVL_Bridge.aFollowingError[6]
    xB39 : BOOL; // GVL_Bridge.aFollowingError[6] >= 2
    rV40 : REAL; // GVL_Hmi.rOverride
    rV41 : REAL; // GVL_Bridge.iWorstJoint
    rV42 : REAL; // GVL_Bridge.stVision.usiClass
    rV43 : REAL; // GVL_Bridge.stVision.rConfidence
    rV44 : REAL; // GVL_Bridge.stVision.lrX
END_VAR

IF GVL_HmiView.xAborted THEN iMachine := 1; ELSIF GVL_HmiView.xHeld THEN iMachine := 2; ELSIF GVL_HmiView.xActing THEN iMachine := 3; ELSIF GVL_HmiView.xManual THEN iMachine := 4; ELSIF GVL_HmiView.xExecute THEN iMachine := 5; ELSIF GVL_HmiView.xIdle THEN iMachine := 6; ELSE iMachine := 0; END_IF
sV1 := TO_STRING(GVL_HmiView.sState);
sV2 := TO_STRING(GVL_HmiView.sMode);
rV3 := ANY_TO_REAL(GVL_HmiView.uiPlaced);
rV4 := ANY_TO_REAL(GVL_Bridge.aJointPosSp[1]);
iP5 := REAL_TO_INT(LIMIT(0.0, (ANY_TO_REAL(GVL_Bridge.aJointPosSp[1]) - (-180.0)) / (360.0), 1.0) * 80.0);
rV6 := ANY_TO_REAL(GVL_Bridge.aJointPosSp[2]);
iP7 := REAL_TO_INT(LIMIT(0.0, (ANY_TO_REAL(GVL_Bridge.aJointPosSp[2]) - (-180.0)) / (360.0), 1.0) * 80.0);
rV8 := ANY_TO_REAL(GVL_Bridge.aJointPosSp[3]);
iP9 := REAL_TO_INT(LIMIT(0.0, (ANY_TO_REAL(GVL_Bridge.aJointPosSp[3]) - (-180.0)) / (360.0), 1.0) * 80.0);
rV10 := ANY_TO_REAL(GVL_Bridge.aJointPosSp[4]);
iP11 := REAL_TO_INT(LIMIT(0.0, (ANY_TO_REAL(GVL_Bridge.aJointPosSp[4]) - (-360.0)) / (720.0), 1.0) * 80.0);
rV12 := ANY_TO_REAL(GVL_Bridge.aJointPosSp[5]);
iP13 := REAL_TO_INT(LIMIT(0.0, (ANY_TO_REAL(GVL_Bridge.aJointPosSp[5]) - (-180.0)) / (360.0), 1.0) * 80.0);
rV14 := ANY_TO_REAL(GVL_Bridge.aJointPosSp[6]);
iP15 := REAL_TO_INT(LIMIT(0.0, (ANY_TO_REAL(GVL_Bridge.aJointPosSp[6]) - (-360.0)) / (720.0), 1.0) * 80.0);
rV16 := ANY_TO_REAL(GVL_Bridge.aFollowingError[1]);
xB17 := ANY_TO_REAL(GVL_Bridge.aFollowingError[1]) >= 2.0;
iP18 := REAL_TO_INT(LIMIT(0.0, (ANY_TO_REAL(GVL_Bridge.aFollowingError[1]) - (0.0)) / (6.0), 1.0) * 80.0);
xB19 := ANY_TO_REAL(GVL_Bridge.aFollowingError[1]) >= 2.0;
rV20 := ANY_TO_REAL(GVL_Bridge.aFollowingError[2]);
xB21 := ANY_TO_REAL(GVL_Bridge.aFollowingError[2]) >= 2.0;
iP22 := REAL_TO_INT(LIMIT(0.0, (ANY_TO_REAL(GVL_Bridge.aFollowingError[2]) - (0.0)) / (6.0), 1.0) * 80.0);
xB23 := ANY_TO_REAL(GVL_Bridge.aFollowingError[2]) >= 2.0;
rV24 := ANY_TO_REAL(GVL_Bridge.aFollowingError[3]);
xB25 := ANY_TO_REAL(GVL_Bridge.aFollowingError[3]) >= 2.0;
iP26 := REAL_TO_INT(LIMIT(0.0, (ANY_TO_REAL(GVL_Bridge.aFollowingError[3]) - (0.0)) / (6.0), 1.0) * 80.0);
xB27 := ANY_TO_REAL(GVL_Bridge.aFollowingError[3]) >= 2.0;
rV28 := ANY_TO_REAL(GVL_Bridge.aFollowingError[4]);
xB29 := ANY_TO_REAL(GVL_Bridge.aFollowingError[4]) >= 2.0;
iP30 := REAL_TO_INT(LIMIT(0.0, (ANY_TO_REAL(GVL_Bridge.aFollowingError[4]) - (0.0)) / (6.0), 1.0) * 80.0);
xB31 := ANY_TO_REAL(GVL_Bridge.aFollowingError[4]) >= 2.0;
rV32 := ANY_TO_REAL(GVL_Bridge.aFollowingError[5]);
xB33 := ANY_TO_REAL(GVL_Bridge.aFollowingError[5]) >= 2.0;
iP34 := REAL_TO_INT(LIMIT(0.0, (ANY_TO_REAL(GVL_Bridge.aFollowingError[5]) - (0.0)) / (6.0), 1.0) * 80.0);
xB35 := ANY_TO_REAL(GVL_Bridge.aFollowingError[5]) >= 2.0;
rV36 := ANY_TO_REAL(GVL_Bridge.aFollowingError[6]);
xB37 := ANY_TO_REAL(GVL_Bridge.aFollowingError[6]) >= 2.0;
iP38 := REAL_TO_INT(LIMIT(0.0, (ANY_TO_REAL(GVL_Bridge.aFollowingError[6]) - (0.0)) / (6.0), 1.0) * 80.0);
xB39 := ANY_TO_REAL(GVL_Bridge.aFollowingError[6]) >= 2.0;
rV40 := ANY_TO_REAL(GVL_Hmi.rOverride);
rV41 := ANY_TO_REAL(GVL_Bridge.iWorstJoint);
rV42 := ANY_TO_REAL(GVL_Bridge.stVision.usiClass);
rV43 := ANY_TO_REAL(GVL_Bridge.stVision.rConfidence);
rV44 := ANY_TO_REAL(GVL_Bridge.stVision.lrX);

END_PROGRAM

// Device/Application/PRG_HMI_Overview
PROGRAM PRG_HMI_Overview
// Generated by codesys-mcp-toolkit for the HMI screen 'Overview' (49 variables). Rebuilt on every export.
VAR
    iMachine : INT; // the machine's state: 0 idle, 1.. the states in order
    sV1 : STRING(80); // GVL_HmiView.sState
    sV2 : STRING(80); // GVL_HmiView.sMode
    rV3 : REAL; // GVL_HmiView.uiPlaced
    rV4 : REAL; // GVL_Bridge.lrBeltVel
    rV5 : REAL; // GVL_HmiView.uiPlaced
    rV6 : REAL; // GVL_Bridge.lrBeltVel
    iP7 : INT; // GVL_Bridge.lrBeltVel
    rV8 : REAL; // GVL_HmiView.uiPlaced
    rV9 : REAL; // PRG_Main.fbCell.aBins[0].uiCount
    xB10 : BOOL; // PRG_Main.fbCell.aBins[0].uiCount >= 27
    iP11 : INT; // PRG_Main.fbCell.aBins[0].uiCount
    xB12 : BOOL; // PRG_Main.fbCell.aBins[0].uiCount >= 27
    rV13 : REAL; // PRG_Main.fbCell.aBins[1].uiCount
    xB14 : BOOL; // PRG_Main.fbCell.aBins[1].uiCount >= 27
    iP15 : INT; // PRG_Main.fbCell.aBins[1].uiCount
    xB16 : BOOL; // PRG_Main.fbCell.aBins[1].uiCount >= 27
    rV17 : REAL; // PRG_Main.fbCell.aBins[2].uiCount
    xB18 : BOOL; // PRG_Main.fbCell.aBins[2].uiCount >= 27
    iP19 : INT; // PRG_Main.fbCell.aBins[2].uiCount
    xB20 : BOOL; // PRG_Main.fbCell.aBins[2].uiCount >= 27
    rV21 : REAL; // PRG_Main.fbCell.aBins[3].uiCount
    xB22 : BOOL; // PRG_Main.fbCell.aBins[3].uiCount >= 27
    iP23 : INT; // PRG_Main.fbCell.aBins[3].uiCount
    xB24 : BOOL; // PRG_Main.fbCell.aBins[3].uiCount >= 27
    rV25 : REAL; // PRG_Main.fbCell.aBins[4].uiCount
    xB26 : BOOL; // PRG_Main.fbCell.aBins[4].uiCount >= 27
    iP27 : INT; // PRG_Main.fbCell.aBins[4].uiCount
    xB28 : BOOL; // PRG_Main.fbCell.aBins[4].uiCount >= 27
    rV29 : REAL; // PRG_Main.fbCell.aBins[5].uiCount
    xB30 : BOOL; // PRG_Main.fbCell.aBins[5].uiCount >= 27
    iP31 : INT; // PRG_Main.fbCell.aBins[5].uiCount
    xB32 : BOOL; // PRG_Main.fbCell.aBins[5].uiCount >= 27
END_VAR

IF GVL_HmiView.xAborted THEN iMachine := 1; ELSIF GVL_HmiView.xHeld THEN iMachine := 2; ELSIF GVL_HmiView.xActing THEN iMachine := 3; ELSIF GVL_HmiView.xManual THEN iMachine := 4; ELSIF GVL_HmiView.xExecute THEN iMachine := 5; ELSIF GVL_HmiView.xIdle THEN iMachine := 6; ELSE iMachine := 0; END_IF
sV1 := TO_STRING(GVL_HmiView.sState);
sV2 := TO_STRING(GVL_HmiView.sMode);
rV3 := ANY_TO_REAL(GVL_HmiView.uiPlaced);
rV4 := ANY_TO_REAL(GVL_Bridge.lrBeltVel);
rV5 := ANY_TO_REAL(GVL_HmiView.uiPlaced);
rV6 := ANY_TO_REAL(GVL_Bridge.lrBeltVel);
iP7 := REAL_TO_INT(LIMIT(0.0, (ANY_TO_REAL(GVL_Bridge.lrBeltVel) - (0.0)) / (150.0), 1.0) * 374.0);
rV8 := ANY_TO_REAL(GVL_HmiView.uiPlaced);
rV9 := ANY_TO_REAL(PRG_Main.fbCell.aBins[0].uiCount);
xB10 := ANY_TO_REAL(PRG_Main.fbCell.aBins[0].uiCount) >= 27.0;
iP11 := REAL_TO_INT(LIMIT(0.0, (ANY_TO_REAL(PRG_Main.fbCell.aBins[0].uiCount) - (0.0)) / (30.0), 1.0) * 80.0);
xB12 := ANY_TO_REAL(PRG_Main.fbCell.aBins[0].uiCount) >= 27.0;
rV13 := ANY_TO_REAL(PRG_Main.fbCell.aBins[1].uiCount);
xB14 := ANY_TO_REAL(PRG_Main.fbCell.aBins[1].uiCount) >= 27.0;
iP15 := REAL_TO_INT(LIMIT(0.0, (ANY_TO_REAL(PRG_Main.fbCell.aBins[1].uiCount) - (0.0)) / (30.0), 1.0) * 80.0);
xB16 := ANY_TO_REAL(PRG_Main.fbCell.aBins[1].uiCount) >= 27.0;
rV17 := ANY_TO_REAL(PRG_Main.fbCell.aBins[2].uiCount);
xB18 := ANY_TO_REAL(PRG_Main.fbCell.aBins[2].uiCount) >= 27.0;
iP19 := REAL_TO_INT(LIMIT(0.0, (ANY_TO_REAL(PRG_Main.fbCell.aBins[2].uiCount) - (0.0)) / (30.0), 1.0) * 80.0);
xB20 := ANY_TO_REAL(PRG_Main.fbCell.aBins[2].uiCount) >= 27.0;
rV21 := ANY_TO_REAL(PRG_Main.fbCell.aBins[3].uiCount);
xB22 := ANY_TO_REAL(PRG_Main.fbCell.aBins[3].uiCount) >= 27.0;
iP23 := REAL_TO_INT(LIMIT(0.0, (ANY_TO_REAL(PRG_Main.fbCell.aBins[3].uiCount) - (0.0)) / (30.0), 1.0) * 80.0);
xB24 := ANY_TO_REAL(PRG_Main.fbCell.aBins[3].uiCount) >= 27.0;
rV25 := ANY_TO_REAL(PRG_Main.fbCell.aBins[4].uiCount);
xB26 := ANY_TO_REAL(PRG_Main.fbCell.aBins[4].uiCount) >= 27.0;
iP27 := REAL_TO_INT(LIMIT(0.0, (ANY_TO_REAL(PRG_Main.fbCell.aBins[4].uiCount) - (0.0)) / (30.0), 1.0) * 80.0);
xB28 := ANY_TO_REAL(PRG_Main.fbCell.aBins[4].uiCount) >= 27.0;
rV29 := ANY_TO_REAL(PRG_Main.fbCell.aBins[5].uiCount);
xB30 := ANY_TO_REAL(PRG_Main.fbCell.aBins[5].uiCount) >= 27.0;
iP31 := REAL_TO_INT(LIMIT(0.0, (ANY_TO_REAL(PRG_Main.fbCell.aBins[5].uiCount) - (0.0)) / (30.0), 1.0) * 80.0);
xB32 := ANY_TO_REAL(PRG_Main.fbCell.aBins[5].uiCount) >= 27.0;

END_PROGRAM

// Device/Application/Visu_Overview
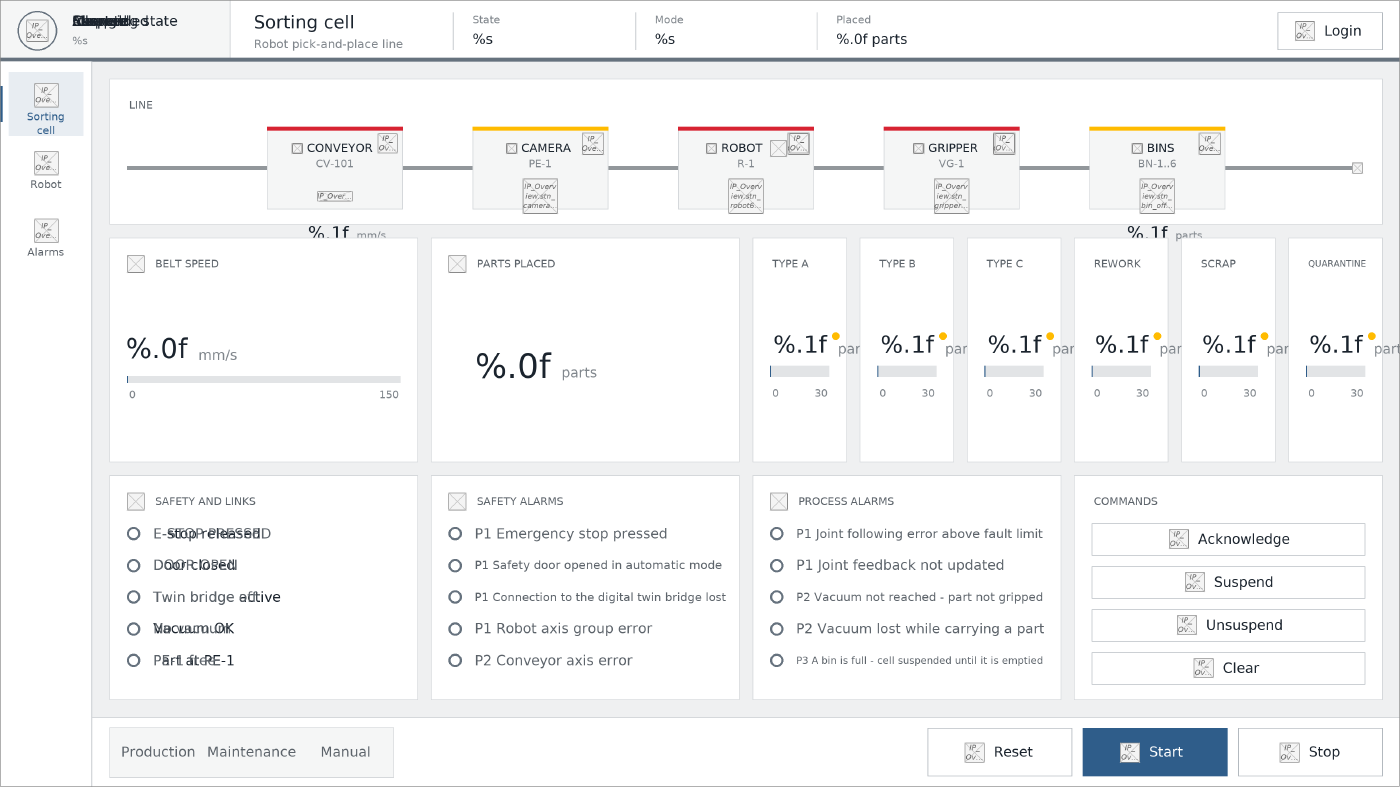
VISUALIZATION Visu_Overview  // 1920x1080
    Rectangle (0,0 1920x84)
    Rectangle (0,83 1920x1)
    Rectangle (0,0 315x83)
    Rectangle (315,0 1x83)
    Rectangle (0,79 1920x5), invisible if: PRG_HMI_Overview.iMachine <> 0
    Ellipse (24,15 54x54), invisible if: PRG_HMI_Overview.iMachine <> 0
    Image (36,27 30x30), invisible if: PRG_HMI_Overview.iMachine <> 0, image: IP_Overview.ic_stop_30_66727e
    Rectangle (96,14 198x30), "Stopped", invisible if: PRG_HMI_Overview.iMachine <> 0
    Rectangle (0,79 1920x5), invisible if: PRG_HMI_Overview.iMachine <> 1
    Ellipse (24,15 54x54), invisible if: PRG_HMI_Overview.iMachine <> 1
    Image (36,27 30x30), invisible if: PRG_HMI_Overview.iMachine <> 1, image: IP_Overview.ic_fault_30_d72332
    Rectangle (96,14 198x30), "Aborted", invisible if: PRG_HMI_Overview.iMachine <> 1
    Rectangle (0,79 1920x5), invisible if: PRG_HMI_Overview.iMachine <> 2
    Ellipse (24,15 54x54), invisible if: PRG_HMI_Overview.iMachine <> 2
    Image (36,27 30x30), invisible if: PRG_HMI_Overview.iMachine <> 2, image: IP_Overview.ic_pause_30_ffbb00
    Rectangle (96,14 198x30), "Suspended", invisible if: PRG_HMI_Overview.iMachine <> 2
    Rectangle (0,79 1920x5), invisible if: PRG_HMI_Overview.iMachine <> 3
    Ellipse (24,15 54x54), invisible if: PRG_HMI_Overview.iMachine <> 3
    Image (36,27 30x30), invisible if: PRG_HMI_Overview.iMachine <> 3, image: IP_Overview.ic_warning_30_ffbb00
    Rectangle (96,14 198x30), "Changing state", invisible if: PRG_HMI_Overview.iMachine <> 3
    Rectangle (0,79 1920x5), invisible if: PRG_HMI_Overview.iMachine <> 4
    Ellipse (24,15 54x54), invisible if: PRG_HMI_Overview.iMachine <> 4
    Image (36,27 30x30), invisible if: PRG_HMI_Overview.iMachine <> 4, image: IP_Overview.ic_manual_30_2f5d8a
    Rectangle (96,14 198x30), "Manual", invisible if: PRG_HMI_Overview.iMachine <> 4
    Rectangle (0,79 1920x5), invisible if: PRG_HMI_Overview.iMachine <> 5
    Ellipse (24,15 54x54), invisible if: PRG_HMI_Overview.iMachine <> 5
    Image (36,27 30x30), invisible if: PRG_HMI_Overview.iMachine <> 5, image: IP_Overview.ic_play_30_66727e
    Rectangle (96,14 198x30), "Execute", invisible if: PRG_HMI_Overview.iMachine <> 5
    Rectangle (0,79 1920x5), invisible if: PRG_HMI_Overview.iMachine <> 6
    Ellipse (24,15 54x54), invisible if: PRG_HMI_Overview.iMachine <> 6
    Image (36,27 30x30), invisible if: PRG_HMI_Overview.iMachine <> 6, image: IP_Overview.ic_stop_30_66727e
    Rectangle (96,14 198x30), "Idle", invisible if: PRG_HMI_Overview.iMachine <> 6
    Rectangle (96,44 198x24), "%s", text variable: GVL_HmiView.sPickStep
    Rectangle (345,11 246x39), "Sorting cell"
    Rectangle (345,47 246x27), "Robot pick-and-place line"
    Rectangle (621,17 1x51)
    Rectangle (645,15 226x24), "State"
    Rectangle (645,39 226x30), "%s", text variable: PRG_HMI_Overview.sV1
    Rectangle (871,17 1x51)
    Rectangle (895,15 226x24), "Mode"
    Rectangle (895,39 226x30), "%s", text variable: PRG_HMI_Overview.sV2
    Rectangle (1120,17 1x51)
    Rectangle (1144,15 163x24), "Placed"
    Rectangle (1144,39 163x30), "%.0f parts", text variable: PRG_HMI_Overview.rV3
    RoundedRectangle (1752,17 144x51)
    Image (1776,29 27x27), image: IP_Overview.ic_login_27_1a232d
    Rectangle (1813,17 81x51), "Login"
    Rectangle (1752,17 144x51)
        OnMouseClick:  Type=Login, OpenCentered=True
    Rectangle (126,984 1794x96)
    Rectangle (126,984 1794x1)
    RoundedRectangle (150,998 390x69)
    RoundedRectangle (155,1002 124x60), colour toggle: GVL_HmiPanel.iModeSelect = 1
    Rectangle (155,1002 124x60), "Production", colour toggle: GVL_HmiPanel.iModeSelect = 1
    Rectangle (155,1002 124x60)
        OnMouseClick: execute { GVL_HmiPanel.iModeSelect := 1; }
    RoundedRectangle (283,1002 124x60), colour toggle: GVL_HmiPanel.iModeSelect = 2
    Rectangle (283,1002 124x60), "Maintenance", colour toggle: GVL_HmiPanel.iModeSelect = 2
    Rectangle (283,1002 124x60)
        OnMouseClick: execute { GVL_HmiPanel.iModeSelect := 2; }
    RoundedRectangle (412,1002 124x60), colour toggle: GVL_HmiPanel.iModeSelect = 3
    Rectangle (412,1002 124x60), "Manual", colour toggle: GVL_HmiPanel.iModeSelect = 3
    Rectangle (412,1002 124x60)
        OnMouseClick: execute { GVL_HmiPanel.iModeSelect := 3; }
    RoundedRectangle (1272,999 198x66), colour toggle: GVL_HmiPanel.xReset
    Image (1323,1019 27x27), image: IP_Overview.ic_reset_27_1a232d
    Rectangle (1360,999 81x66), "Reset"
    Rectangle (1272,999 198x66)
        tap GVL_HmiPanel.xReset
    RoundedRectangle (1485,999 198x66), colour toggle: GVL_HmiPanel.xStart
    Image (1536,1019 27x27), image: IP_Overview.ic_play_27_ffffff
    Rectangle (1573,999 81x66), "Start"
    Rectangle (1485,999 198x66)
        tap GVL_HmiPanel.xStart
    RoundedRectangle (1698,999 198x66), colour toggle: GVL_HmiPanel.xStop
    Image (1755,1019 27x27), image: IP_Overview.ic_stop_27_1a232d
    Rectangle (1792,999 69x66), "Stop"
    Rectangle (1698,999 198x66)
        tap GVL_HmiPanel.xStop
    Rectangle (0,84 126x996)
    Rectangle (125,84 1x996)
    RoundedRectangle (12,99 102x87)
    RoundedRectangle (0,118 3x49)
    Image (47,114 33x33), image: IP_Overview.ic_home_33_2f5d8a
    Rectangle (15,150 96x20), "Sorting"
    Rectangle (15,169 96x20), "cell"
    Image (47,207 33x33), image: IP_Overview.ic_machine_33_5c636a
    Rectangle (15,243 96x20), "Robot"
    Rectangle (12,192 102x87)
        OnMouseClick:  Assign=Visu_Robot, Type=Assignment
    Image (47,300 33x33), image: IP_Overview.ic_alarm_33_5c636a
    Rectangle (15,336 96x20), "Alarms"
    Rectangle (12,285 102x87)
        OnMouseClick:  Assign=Visu_Alarms, Type=Assignment
    RoundedRectangle (150,108 1746x200)
    Rectangle (174,129 1698x30), "LINE"
    Rectangle (174,228 1683x5)
    Image (1854,223 15x15), image: IP_Overview.arrow_r_15_92979b
    RoundedRectangle (366,174 186x113)
    Rectangle (366,174 186x5)
    Rectangle (366,174 186x5), invisible if: NOT (GVL_HmiView.axAlarmActive[5])
    Image (400,196 15x15), invisible if: NOT (GVL_HmiView.xBeltRunning), image: IP_Overview.sign_run_15
    Image (401,197 13x13), invisible if: GVL_HmiView.xBeltRunning, image: IP_Overview.sign_stop_13
    Rectangle (418,191 110x24), "CONVEYOR"
    Rectangle (372,214 174x21), "CV-101"
    Image (435,262 48x14), image: IP_Overview.stn_conveyor_off_48x14
        p84334746: SEL(GVL_HmiView.xBeltRunning, 'IP_Overview.stn_conveyor_off_48x14', 'IP_Overview.stn_conveyor_on_48x14')
    Rectangle (362,302 119x36), "%.1f", text variable: PRG_HMI_Overview.rV4
    Rectangle (486,311 74x24), "mm/s"
    Image (518,183 27x27), invisible if: NOT (GVL_HmiView.axAlarmActive[5]), image: IP_Overview.sign_alarm_27
    Rectangle (366,174 186x113)
        OnMouseClick:  Assign=Visu_Robot, Type=Assignment
    RoundedRectangle (648,174 186x113)
    Rectangle (648,174 186x5)
    Rectangle (648,174 186x5), invisible if: NOT (GVL_HmiView.axAlarm[13])
    Image (694,196 15x15), invisible if: NOT (GVL_Bridge.xPE1), image: IP_Overview.sign_run_15
    Image (695,197 13x13), invisible if: GVL_Bridge.xPE1, image: IP_Overview.sign_stop_13
    Rectangle (712,191 85x24), "CAMERA"
    Rectangle (654,214 174x21), "PE-1"
    Image (717,245 48x48), image: IP_Overview.stn_camera_off_48x48
        p84334746: SEL(GVL_Bridge.xPE1, 'IP_Overview.stn_camera_off_48x48', 'IP_Overview.stn_camera_on_48x48')
    Image (798,182 30x30), invisible if: NOT (GVL_HmiView.axAlarm[13]), image: IP_Overview.sign_warning_30
    Rectangle (648,174 186x113)
        OnMouseClick:  Assign=Visu_Alarms, Type=Assignment
    RoundedRectangle (930,174 186x113)
    Rectangle (930,174 186x5)
    Rectangle (930,174 186x5), invisible if: NOT (GVL_HmiView.axAlarmActive[6])
    Rectangle (930,174 186x5), invisible if: NOT (GVL_HmiView.axAlarmActive[4])
    Image (968,196 15x15), invisible if: NOT (GVL_HmiView.xRobotMoving), image: IP_Overview.sign_run_15
    Image (969,197 13x13), invisible if: GVL_HmiView.xRobotMoving, image: IP_Overview.sign_stop_13
    Rectangle (986,191 73x24), "ROBOT"
    Image (1056,192 23x23), invisible if: NOT (GVL_HmiView.xManual), image: IP_Overview.ic_manual_23_2f5d8a
    Rectangle (936,214 174x21), "R-1"
    Image (999,245 48x48), image: IP_Overview.stn_robot6_off_48x48
        p84334746: SEL(GVL_HmiView.xRobotMoving, 'IP_Overview.stn_robot6_off_48x48', 'IP_Overview.stn_robot6_on_48x48')
    Image (1080,182 30x30), invisible if: NOT ((GVL_HmiView.axAlarmActive[6]) AND NOT (GVL_HmiView.axAlarmActive[4])), image: IP_Overview.sign_warning_30
    Image (1082,183 27x27), invisible if: NOT (GVL_HmiView.axAlarmActive[4]), image: IP_Overview.sign_alarm_27
    Rectangle (930,174 186x113)
        OnMouseClick:  Assign=Visu_Robot, Type=Assignment
    RoundedRectangle (1212,174 186x113)
    Rectangle (1212,174 186x5)
    Rectangle (1212,174 186x5), invisible if: NOT (GVL_HmiView.axAlarm[9])
    Rectangle (1212,174 186x5), invisible if: NOT (GVL_HmiView.axAlarm[10])
    Image (1252,196 15x15), invisible if: NOT (GVL_Bridge.xVacuumOn), image: IP_Overview.sign_run_15
    Image (1253,197 13x13), invisible if: GVL_Bridge.xVacuumOn, image: IP_Overview.sign_stop_13
    Rectangle (1270,191 98x24), "GRIPPER"
    Rectangle (1218,214 174x21), "VG-1"
    Image (1281,245 48x48), image: IP_Overview.stn_gripper_off_48x48
        p84334746: SEL(GVL_Bridge.xVacuumOn, 'IP_Overview.stn_gripper_off_48x48', 'IP_Overview.stn_gripper_on_48x48')
    Image (1362,182 30x30), invisible if: NOT ((GVL_HmiView.axAlarm[9]) AND NOT (GVL_HmiView.axAlarm[10])), image: IP_Overview.sign_warning_30
    Image (1364,183 27x27), invisible if: NOT (GVL_HmiView.axAlarm[10]), image: IP_Overview.sign_alarm_27
    Rectangle (1212,174 186x113)
        OnMouseClick:  Assign=Visu_Robot, Type=Assignment
    RoundedRectangle (1494,174 186x113)
    Rectangle (1494,174 186x5)
    Rectangle (1494,174 186x5), invisible if: NOT (GVL_HmiView.xAnyBinFull)
    Image (1552,196 15x15), invisible if: NOT (GVL_HmiView.xExecute), image: IP_Overview.sign_run_15
    Image (1553,197 13x13), invisible if: GVL_HmiView.xExecute, image: IP_Overview.sign_stop_13
    Rectangle (1570,191 61x24), "BINS"
    Rectangle (1500,214 174x21), "BN-1..6"
    Image (1563,245 48x48), image: IP_Overview.stn_bin_off_48x48
        p84334746: SEL(GVL_HmiView.xExecute, 'IP_Overview.stn_bin_off_48x48', 'IP_Overview.stn_bin_on_48x48')
    Rectangle (1485,302 119x36), "%.1f", text variable: PRG_HMI_Overview.rV5
    Rectangle (1609,311 84x24), "parts"
    Image (1644,182 30x30), invisible if: NOT (GVL_HmiView.xAnyBinFull), image: IP_Overview.sign_warning_30
    Rectangle (1494,174 186x113)
        OnMouseClick:  Assign=Visu_Alarms, Type=Assignment
    RoundedRectangle (150,326 423x308)
    Image (174,350 24x24), image: IP_Overview.ic_speed_24_80868c
    Rectangle (210,347 339x30), "BELT SPEED"
    Rectangle (174,445 86x66), "%.0f", text variable: PRG_HMI_Overview.rV6
    Rectangle (269,469 135x37), "mm/s"
    RoundedRectangle (174,516 375x9)
    RoundedRectangle (174,516 1x9)
        p874137650: PRG_HMI_Overview.iP7
    Rectangle (174,531 188x21), "0"
    Rectangle (362,531 188x21), "150"
    RoundedRectangle (591,326 423x308)
    Image (615,350 24x24), image: IP_Overview.ic_count_24_80868c
    Rectangle (651,347 339x30), "PARTS PLACED"
    Rectangle (615,469 143x66), "%.0f", text variable: PRG_HMI_Overview.rV8
    Rectangle (767,493 135x37), "parts"
    RoundedRectangle (1032,326 129x308)
    Rectangle (1056,347 81x30), "TYPE A"
    Rectangle (1056,449 81x47), "%.1f", text variable: PRG_HMI_Overview.rV9
    Ellipse (1141,456 10x10), invisible if: NOT PRG_HMI_Overview.xB10
    Rectangle (1146,466 135x26), "parts"
    RoundedRectangle (1056,502 81x15)
    RoundedRectangle (1056,502 1x15), colour toggle: PRG_HMI_Overview.xB12
        p874137650: PRG_HMI_Overview.iP11
    Rectangle (1056,529 41x21), "0"
    Rectangle (1097,529 41x21), "30"
    RoundedRectangle (1179,326 129x308)
    Rectangle (1203,347 81x30), "TYPE B"
    Rectangle (1203,449 81x47), "%.1f", text variable: PRG_HMI_Overview.rV13
    Ellipse (1288,456 10x10), invisible if: NOT PRG_HMI_Overview.xB14
    Rectangle (1293,466 135x26), "parts"
    RoundedRectangle (1203,502 81x15)
    RoundedRectangle (1203,502 1x15), colour toggle: PRG_HMI_Overview.xB16
        p874137650: PRG_HMI_Overview.iP15
    Rectangle (1203,529 41x21), "0"
    Rectangle (1244,529 41x21), "30"
    RoundedRectangle (1326,326 129x308)
    Rectangle (1350,347 81x30), "TYPE C"
    Rectangle (1350,449 81x47), "%.1f", text variable: PRG_HMI_Overview.rV17
    Ellipse (1435,456 10x10), invisible if: NOT PRG_HMI_Overview.xB18
    Rectangle (1440,466 135x26), "parts"
    RoundedRectangle (1350,502 81x15)
    RoundedRectangle (1350,502 1x15), colour toggle: PRG_HMI_Overview.xB20
        p874137650: PRG_HMI_Overview.iP19
    Rectangle (1350,529 41x21), "0"
    Rectangle (1391,529 41x21), "30"
    RoundedRectangle (1473,326 129x308)
    Rectangle (1497,347 81x30), "REWORK"
    Rectangle (1497,449 81x47), "%.1f", text variable: PRG_HMI_Overview.rV21
    Ellipse (1582,456 10x10), invisible if: NOT PRG_HMI_Overview.xB22
    Rectangle (1587,466 135x26), "parts"
    RoundedRectangle (1497,502 81x15)
    RoundedRectangle (1497,502 1x15), colour toggle: PRG_HMI_Overview.xB24
        p874137650: PRG_HMI_Overview.iP23
    Rectangle (1497,529 41x21), "0"
    Rectangle (1538,529 41x21), "30"
    RoundedRectangle (1620,326 129x308)
    Rectangle (1644,347 81x30), "SCRAP"
    Rectangle (1644,449 81x47), "%.1f", text variable: PRG_HMI_Overview.rV25
    Ellipse (1729,456 10x10), invisible if: NOT PRG_HMI_Overview.xB26
    Rectangle (1734,466 135x26), "parts"
    RoundedRectangle (1644,502 81x15)
    RoundedRectangle (1644,502 1x15), colour toggle: PRG_HMI_Overview.xB28
        p874137650: PRG_HMI_Overview.iP27
    Rectangle (1644,529 41x21), "0"
    Rectangle (1685,529 41x21), "30"
    RoundedRectangle (1767,326 129x308)
    Rectangle (1791,347 81x30), "QUARANTINE"
    Rectangle (1791,449 81x47), "%.1f", text variable: PRG_HMI_Overview.rV29
    Ellipse (1876,456 10x10), invisible if: NOT PRG_HMI_Overview.xB30
    Rectangle (1881,466 135x26), "parts"
    RoundedRectangle (1791,502 81x15)
    RoundedRectangle (1791,502 1x15), colour toggle: PRG_HMI_Overview.xB32
        p874137650: PRG_HMI_Overview.iP31
    Rectangle (1791,529 41x21), "0"
    Rectangle (1832,529 41x21), "30"
    RoundedRectangle (150,652 423x308)
    Image (174,676 24x24), image: IP_Overview.ic_info_24_80868c
    Rectangle (210,673 339x30), "SAFETY AND LINKS"
    Ellipse (174,723 18x18), colour toggle: GVL_Bridge.xEStopOk
    Rectangle (207,718 342x29), "E-stop released", invisible if: NOT (GVL_Bridge.xEStopOk)
    Rectangle (207,718 342x29), "E-STOP PRESSED", invisible if: GVL_Bridge.xEStopOk
    Ellipse (174,767 18x18), colour toggle: GVL_Bridge.xDoorClosed
    Rectangle (207,761 342x29), "Door closed", invisible if: NOT (GVL_Bridge.xDoorClosed)
    Rectangle (207,761 342x29), "DOOR OPEN", invisible if: GVL_Bridge.xDoorClosed
    Ellipse (174,810 18x18), colour toggle: GVL_Bridge.xTwinActive
    Rectangle (207,805 342x29), "Twin bridge active", invisible if: NOT (GVL_Bridge.xTwinActive)
    Rectangle (207,805 342x29), "Twin bridge off", invisible if: GVL_Bridge.xTwinActive
    Ellipse (174,854 18x18), colour toggle: GVL_Bridge.xVacuumOk
    Rectangle (207,848 342x29), "Vacuum OK", invisible if: NOT (GVL_Bridge.xVacuumOk)
    Rectangle (207,848 342x29), "No vacuum", invisible if: GVL_Bridge.xVacuumOk
    Ellipse (174,897 18x18), colour toggle: GVL_Bridge.xPE1
    Rectangle (207,892 342x29), "Part at PE-1", invisible if: NOT (GVL_Bridge.xPE1)
    Rectangle (207,892 342x29), "PE-1 free", invisible if: GVL_Bridge.xPE1
    RoundedRectangle (591,652 423x308)
    Image (615,676 24x24), image: IP_Overview.ic_alarm_24_80868c
    Rectangle (651,673 339x30), "SAFETY ALARMS"
    Ellipse (615,723 18x18), colour toggle: GVL_HmiView.axAlarm[1]
    Rectangle (648,718 342x29), "P1 Emergency stop pressed", colour toggle: GVL_HmiView.axAlarm[1]
    Ellipse (615,767 18x18), colour toggle: GVL_HmiView.axAlarm[2]
    Rectangle (648,761 342x29), "P1 Safety door opened in automatic mode", colour toggle: GVL_HmiView.axAlarm[2]
    Ellipse (615,810 18x18), colour toggle: GVL_HmiView.axAlarm[3]
    Rectangle (648,805 342x29), "P1 Connection to the digital twin bridge lost", colour toggle: GVL_HmiView.axAlarm[3]
    Ellipse (615,854 18x18), colour toggle: GVL_HmiView.axAlarm[4]
    Rectangle (648,848 342x29), "P1 Robot axis group error", colour toggle: GVL_HmiView.axAlarm[4]
    Ellipse (615,897 18x18), colour toggle: GVL_HmiView.axAlarm[5]
    Rectangle (648,892 342x29), "P2 Conveyor axis error", colour toggle: GVL_HmiView.axAlarm[5]
    RoundedRectangle (1032,652 423x308)
    Image (1056,676 24x24), image: IP_Overview.ic_alarm_24_80868c
    Rectangle (1092,673 339x30), "PROCESS ALARMS"
    Ellipse (1056,723 18x18), colour toggle: GVL_HmiView.axAlarm[7]
    Rectangle (1089,718 342x29), "P1 Joint following error above fault limit", colour toggle: GVL_HmiView.axAlarm[7]
    Ellipse (1056,767 18x18), colour toggle: GVL_HmiView.axAlarm[8]
    Rectangle (1089,761 342x29), "P1 Joint feedback not updated", colour toggle: GVL_HmiView.axAlarm[8]
    Ellipse (1056,810 18x18), colour toggle: GVL_HmiView.axAlarm[9]
    Rectangle (1089,805 342x29), "P2 Vacuum not reached - part not gripped", colour toggle: GVL_HmiView.axAlarm[9]
    Ellipse (1056,854 18x18), colour toggle: GVL_HmiView.axAlarm[10]
    Rectangle (1089,848 342x29), "P2 Vacuum lost while carrying a part", colour toggle: GVL_HmiView.axAlarm[10]
    Ellipse (1056,897 18x18), colour toggle: GVL_HmiView.axAlarm[12]
    Rectangle (1089,892 342x29), "P3 A bin is full - cell suspended until it is emptied", colour toggle: GVL_HmiView.axAlarm[12]
    RoundedRectangle (1473,652 423x308)
    Rectangle (1497,673 375x30), "COMMANDS"
    RoundedRectangle (1497,718 375x44), colour toggle: GVL_HmiPanel.xAckAll
    Image (1603,726 27x27), image: IP_Overview.ic_check_27_1a232d
    Rectangle (1640,718 149x44), "Acknowledge"
    Rectangle (1497,718 375x44)
        tap GVL_HmiPanel.xAckAll
    RoundedRectangle (1497,777 375x44), colour toggle: GVL_HmiPanel.xSuspend
    Image (1625,785 27x27), image: IP_Overview.ic_pause_27_1a232d
    Rectangle (1662,777 103x44), "Suspend"
    Rectangle (1497,777 375x44)
        tap GVL_HmiPanel.xSuspend
    RoundedRectangle (1497,836 375x44), colour toggle: GVL_HmiPanel.xUnsuspend
    Image (1614,844 27x27), image: IP_Overview.ic_play_27_1a232d
    Rectangle (1651,836 126x44), "Unsuspend"
    Rectangle (1497,836 375x44)
        tap GVL_HmiPanel.xUnsuspend
    RoundedRectangle (1497,895 375x44), colour toggle: GVL_HmiPanel.xClear
    Image (1637,903 27x27), image: IP_Overview.ic_reset_27_1a232d
    Rectangle (1674,895 81x44), "Clear"
    Rectangle (1497,895 375x44)
        tap GVL_HmiPanel.xClear
END_VISUALIZATION

// Device/Application/Visu_Robot
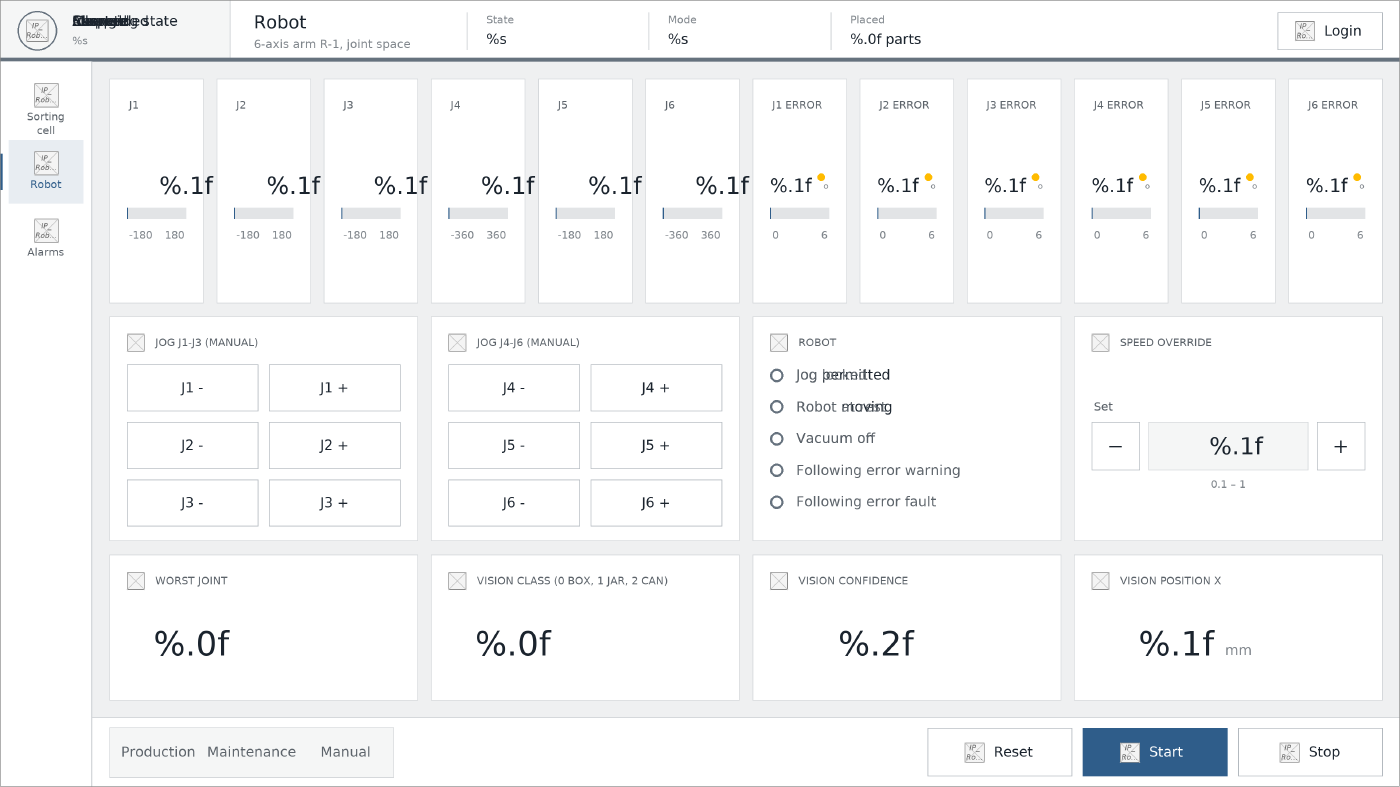
VISUALIZATION Visu_Robot  // 1920x1080
    Rectangle (0,0 1920x84)
    Rectangle (0,83 1920x1)
    Rectangle (0,0 315x83)
    Rectangle (315,0 1x83)
    Rectangle (0,79 1920x5), invisible if: PRG_HMI_Robot.iMachine <> 0
    Ellipse (24,15 54x54), invisible if: PRG_HMI_Robot.iMachine <> 0
    Image (36,27 30x30), invisible if: PRG_HMI_Robot.iMachine <> 0, image: IP_Robot.ic_stop_30_66727e
    Rectangle (96,14 198x30), "Stopped", invisible if: PRG_HMI_Robot.iMachine <> 0
    Rectangle (0,79 1920x5), invisible if: PRG_HMI_Robot.iMachine <> 1
    Ellipse (24,15 54x54), invisible if: PRG_HMI_Robot.iMachine <> 1
    Image (36,27 30x30), invisible if: PRG_HMI_Robot.iMachine <> 1, image: IP_Robot.ic_fault_30_d72332
    Rectangle (96,14 198x30), "Aborted", invisible if: PRG_HMI_Robot.iMachine <> 1
    Rectangle (0,79 1920x5), invisible if: PRG_HMI_Robot.iMachine <> 2
    Ellipse (24,15 54x54), invisible if: PRG_HMI_Robot.iMachine <> 2
    Image (36,27 30x30), invisible if: PRG_HMI_Robot.iMachine <> 2, image: IP_Robot.ic_pause_30_ffbb00
    Rectangle (96,14 198x30), "Suspended", invisible if: PRG_HMI_Robot.iMachine <> 2
    Rectangle (0,79 1920x5), invisible if: PRG_HMI_Robot.iMachine <> 3
    Ellipse (24,15 54x54), invisible if: PRG_HMI_Robot.iMachine <> 3
    Image (36,27 30x30), invisible if: PRG_HMI_Robot.iMachine <> 3, image: IP_Robot.ic_warning_30_ffbb00
    Rectangle (96,14 198x30), "Changing state", invisible if: PRG_HMI_Robot.iMachine <> 3
    Rectangle (0,79 1920x5), invisible if: PRG_HMI_Robot.iMachine <> 4
    Ellipse (24,15 54x54), invisible if: PRG_HMI_Robot.iMachine <> 4
    Image (36,27 30x30), invisible if: PRG_HMI_Robot.iMachine <> 4, image: IP_Robot.ic_manual_30_2f5d8a
    Rectangle (96,14 198x30), "Manual", invisible if: PRG_HMI_Robot.iMachine <> 4
    Rectangle (0,79 1920x5), invisible if: PRG_HMI_Robot.iMachine <> 5
    Ellipse (24,15 54x54), invisible if: PRG_HMI_Robot.iMachine <> 5
    Image (36,27 30x30), invisible if: PRG_HMI_Robot.iMachine <> 5, image: IP_Robot.ic_play_30_66727e
    Rectangle (96,14 198x30), "Execute", invisible if: PRG_HMI_Robot.iMachine <> 5
    Rectangle (0,79 1920x5), invisible if: PRG_HMI_Robot.iMachine <> 6
    Ellipse (24,15 54x54), invisible if: PRG_HMI_Robot.iMachine <> 6
    Image (36,27 30x30), invisible if: PRG_HMI_Robot.iMachine <> 6, image: IP_Robot.ic_stop_30_66727e
    Rectangle (96,14 198x30), "Idle", invisible if: PRG_HMI_Robot.iMachine <> 6
    Rectangle (96,44 198x24), "%s", text variable: GVL_HmiView.sPickStep
    Rectangle (345,11 265x39), "Robot"
    Rectangle (345,47 265x27), "6-axis arm R-1, joint space"
    Rectangle (640,17 1x51)
    Rectangle (664,15 226x24), "State"
    Rectangle (664,39 226x30), "%s", text variable: PRG_HMI_Robot.sV1
    Rectangle (889,17 1x51)
    Rectangle (913,15 226x24), "Mode"
    Rectangle (913,39 226x30), "%s", text variable: PRG_HMI_Robot.sV2
    Rectangle (1139,17 1x51)
    Rectangle (1163,15 163x24), "Placed"
    Rectangle (1163,39 163x30), "%.0f parts", text variable: PRG_HMI_Robot.rV3
    RoundedRectangle (1752,17 144x51)
    Image (1776,29 27x27), image: IP_Robot.ic_login_27_1a232d
    Rectangle (1813,17 81x51), "Login"
    Rectangle (1752,17 144x51)
        OnMouseClick:  Type=Login, OpenCentered=True
    Rectangle (126,984 1794x96)
    Rectangle (126,984 1794x1)
    RoundedRectangle (150,998 390x69)
    RoundedRectangle (155,1002 124x60), colour toggle: GVL_HmiPanel.iModeSelect = 1
    Rectangle (155,1002 124x60), "Production", colour toggle: GVL_HmiPanel.iModeSelect = 1
    Rectangle (155,1002 124x60)
        OnMouseClick: execute { GVL_HmiPanel.iModeSelect := 1; }
    RoundedRectangle (283,1002 124x60), colour toggle: GVL_HmiPanel.iModeSelect = 2
    Rectangle (283,1002 124x60), "Maintenance", colour toggle: GVL_HmiPanel.iModeSelect = 2
    Rectangle (283,1002 124x60)
        OnMouseClick: execute { GVL_HmiPanel.iModeSelect := 2; }
    RoundedRectangle (412,1002 124x60), colour toggle: GVL_HmiPanel.iModeSelect = 3
    Rectangle (412,1002 124x60), "Manual", colour toggle: GVL_HmiPanel.iModeSelect = 3
    Rectangle (412,1002 124x60)
        OnMouseClick: execute { GVL_HmiPanel.iModeSelect := 3; }
    RoundedRectangle (1272,999 198x66), colour toggle: GVL_HmiPanel.xReset
    Image (1323,1019 27x27), image: IP_Robot.ic_reset_27_1a232d
    Rectangle (1360,999 81x66), "Reset"
    Rectangle (1272,999 198x66)
        tap GVL_HmiPanel.xReset
    RoundedRectangle (1485,999 198x66), colour toggle: GVL_HmiPanel.xStart
    Image (1536,1019 27x27), image: IP_Robot.ic_play_27_ffffff
    Rectangle (1573,999 81x66), "Start"
    Rectangle (1485,999 198x66)
        tap GVL_HmiPanel.xStart
    RoundedRectangle (1698,999 198x66), colour toggle: GVL_HmiPanel.xStop
    Image (1755,1019 27x27), image: IP_Robot.ic_stop_27_1a232d
    Rectangle (1792,999 69x66), "Stop"
    Rectangle (1698,999 198x66)
        tap GVL_HmiPanel.xStop
    Rectangle (0,84 126x996)
    Rectangle (125,84 1x996)
    Image (47,114 33x33), image: IP_Robot.ic_home_33_5c636a
    Rectangle (15,150 96x20), "Sorting"
    Rectangle (15,169 96x20), "cell"
    Rectangle (12,99 102x87)
        OnMouseClick:  Assign=Visu_Overview, Type=Assignment
    RoundedRectangle (12,192 102x87)
    RoundedRectangle (0,211 3x49)
    Image (47,207 33x33), image: IP_Robot.ic_machine_33_2f5d8a
    Rectangle (15,243 96x20), "Robot"
    Image (47,300 33x33), image: IP_Robot.ic_alarm_33_5c636a
    Rectangle (15,336 96x20), "Alarms"
    Rectangle (12,285 102x87)
        OnMouseClick:  Assign=Visu_Alarms, Type=Assignment
    RoundedRectangle (150,108 129x308)
    Rectangle (174,129 81x30), "J1"
    Rectangle (174,231 121x47), "%.1f", text variable: PRG_HMI_Robot.rV4
    Rectangle (304,248 135x26), "°"
    RoundedRectangle (174,285 81x15)
    RoundedRectangle (174,285 1x15)
        p874137650: PRG_HMI_Robot.iP5
    Rectangle (174,312 41x21), "-180"
    Rectangle (215,312 41x21), "180"
    RoundedRectangle (297,108 129x308)
    Rectangle (321,129 81x30), "J2"
    Rectangle (321,231 121x47), "%.1f", text variable: PRG_HMI_Robot.rV6
    Rectangle (451,248 135x26), "°"
    RoundedRectangle (321,285 81x15)
    RoundedRectangle (321,285 1x15)
        p874137650: PRG_HMI_Robot.iP7
    Rectangle (321,312 41x21), "-180"
    Rectangle (362,312 41x21), "180"
    RoundedRectangle (444,108 129x308)
    Rectangle (468,129 81x30), "J3"
    Rectangle (468,231 121x47), "%.1f", text variable: PRG_HMI_Robot.rV8
    Rectangle (598,248 135x26), "°"
    RoundedRectangle (468,285 81x15)
    RoundedRectangle (468,285 1x15)
        p874137650: PRG_HMI_Robot.iP9
    Rectangle (468,312 41x21), "-180"
    Rectangle (509,312 41x21), "180"
    RoundedRectangle (591,108 129x308)
    Rectangle (615,129 81x30), "J4"
    Rectangle (615,231 121x47), "%.1f", text variable: PRG_HMI_Robot.rV10
    Rectangle (745,248 135x26), "°"
    RoundedRectangle (615,285 81x15)
    RoundedRectangle (615,285 1x15)
        p874137650: PRG_HMI_Robot.iP11
    Rectangle (615,312 41x21), "-360"
    Rectangle (656,312 41x21), "360"
    RoundedRectangle (738,108 129x308)
    Rectangle (762,129 81x30), "J5"
    Rectangle (762,231 121x47), "%.1f", text variable: PRG_HMI_Robot.rV12
    Rectangle (892,248 135x26), "°"
    RoundedRectangle (762,285 81x15)
    RoundedRectangle (762,285 1x15)
        p874137650: PRG_HMI_Robot.iP13
    Rectangle (762,312 41x21), "-180"
    Rectangle (803,312 41x21), "180"
    RoundedRectangle (885,108 129x308)
    Rectangle (909,129 81x30), "J6"
    Rectangle (909,231 121x47), "%.1f", text variable: PRG_HMI_Robot.rV14
    Rectangle (1039,248 135x26), "°"
    RoundedRectangle (909,285 81x15)
    RoundedRectangle (909,285 1x15)
        p874137650: PRG_HMI_Robot.iP15
    Rectangle (909,312 41x21), "-360"
    Rectangle (950,312 41x21), "360"
    RoundedRectangle (1032,108 129x308)
    Rectangle (1056,129 81x30), "J1 ERROR"
    Rectangle (1056,231 60x47), "%.1f", text variable: PRG_HMI_Robot.rV16
    Ellipse (1121,238 10x10), invisible if: NOT PRG_HMI_Robot.xB17
    Rectangle (1125,248 135x26), "°"
    RoundedRectangle (1056,285 81x15)
    RoundedRectangle (1056,285 1x15), colour toggle: PRG_HMI_Robot.xB19
        p874137650: PRG_HMI_Robot.iP18
    Rectangle (1056,312 41x21), "0"
    Rectangle (1097,312 41x21), "6"
    RoundedRectangle (1179,108 129x308)
    Rectangle (1203,129 81x30), "J2 ERROR"
    Rectangle (1203,231 60x47), "%.1f", text variable: PRG_HMI_Robot.rV20
    Ellipse (1268,238 10x10), invisible if: NOT PRG_HMI_Robot.xB21
    Rectangle (1272,248 135x26), "°"
    RoundedRectangle (1203,285 81x15)
    RoundedRectangle (1203,285 1x15), colour toggle: PRG_HMI_Robot.xB23
        p874137650: PRG_HMI_Robot.iP22
    Rectangle (1203,312 41x21), "0"
    Rectangle (1244,312 41x21), "6"
    RoundedRectangle (1326,108 129x308)
    Rectangle (1350,129 81x30), "J3 ERROR"
    Rectangle (1350,231 60x47), "%.1f", text variable: PRG_HMI_Robot.rV24
    Ellipse (1415,238 10x10), invisible if: NOT PRG_HMI_Robot.xB25
    Rectangle (1419,248 135x26), "°"
    RoundedRectangle (1350,285 81x15)
    RoundedRectangle (1350,285 1x15), colour toggle: PRG_HMI_Robot.xB27
        p874137650: PRG_HMI_Robot.iP26
    Rectangle (1350,312 41x21), "0"
    Rectangle (1391,312 41x21), "6"
    RoundedRectangle (1473,108 129x308)
    Rectangle (1497,129 81x30), "J4 ERROR"
    Rectangle (1497,231 60x47), "%.1f", text variable: PRG_HMI_Robot.rV28
    Ellipse (1562,238 10x10), invisible if: NOT PRG_HMI_Robot.xB29
    Rectangle (1566,248 135x26), "°"
    RoundedRectangle (1497,285 81x15)
    RoundedRectangle (1497,285 1x15), colour toggle: PRG_HMI_Robot.xB31
        p874137650: PRG_HMI_Robot.iP30
    Rectangle (1497,312 41x21), "0"
    Rectangle (1538,312 41x21), "6"
    RoundedRectangle (1620,108 129x308)
    Rectangle (1644,129 81x30), "J5 ERROR"
    Rectangle (1644,231 60x47), "%.1f", text variable: PRG_HMI_Robot.rV32
    Ellipse (1709,238 10x10), invisible if: NOT PRG_HMI_Robot.xB33
    Rectangle (1713,248 135x26), "°"
    RoundedRectangle (1644,285 81x15)
    RoundedRectangle (1644,285 1x15), colour toggle: PRG_HMI_Robot.xB35
        p874137650: PRG_HMI_Robot.iP34
    Rectangle (1644,312 41x21), "0"
    Rectangle (1685,312 41x21), "6"
    RoundedRectangle (1767,108 129x308)
    Rectangle (1791,129 81x30), "J6 ERROR"
    Rectangle (1791,231 60x47), "%.1f", text variable: PRG_HMI_Robot.rV36
    Ellipse (1856,238 10x10), invisible if: NOT PRG_HMI_Robot.xB37
    Rectangle (1860,248 135x26), "°"
    RoundedRectangle (1791,285 81x15)
    RoundedRectangle (1791,285 1x15), colour toggle: PRG_HMI_Robot.xB39
        p874137650: PRG_HMI_Robot.iP38
    Rectangle (1791,312 41x21), "0"
    Rectangle (1832,312 41x21), "6"
    RoundedRectangle (150,434 423x308)
    Image (174,458 24x24), image: IP_Robot.ic_manual_24_80868c
    Rectangle (210,455 339x30), "JOG J1-J3 (MANUAL)"
    RoundedRectangle (174,500 180x64), colour toggle: GVL_Hmi.axJogMinus[1]
    Rectangle (174,500 180x64), "J1 -"
    Rectangle (174,500 180x64)
        tap GVL_Hmi.axJogMinus[1]
    RoundedRectangle (369,500 180x64), colour toggle: GVL_Hmi.axJogPlus[1]
    Rectangle (369,500 180x64), "J1 +"
    Rectangle (369,500 180x64)
        tap GVL_Hmi.axJogPlus[1]
    RoundedRectangle (174,579 180x64), colour toggle: GVL_Hmi.axJogMinus[2]
    Rectangle (174,579 180x64), "J2 -"
    Rectangle (174,579 180x64)
        tap GVL_Hmi.axJogMinus[2]
    RoundedRectangle (369,579 180x64), colour toggle: GVL_Hmi.axJogPlus[2]
    Rectangle (369,579 180x64), "J2 +"
    Rectangle (369,579 180x64)
        tap GVL_Hmi.axJogPlus[2]
    RoundedRectangle (174,658 180x64), colour toggle: GVL_Hmi.axJogMinus[3]
    Rectangle (174,658 180x64), "J3 -"
    Rectangle (174,658 180x64)
        tap GVL_Hmi.axJogMinus[3]
    RoundedRectangle (369,658 180x64), colour toggle: GVL_Hmi.axJogPlus[3]
    Rectangle (369,658 180x64), "J3 +"
    Rectangle (369,658 180x64)
        tap GVL_Hmi.axJogPlus[3]
    RoundedRectangle (591,434 423x308)
    Image (615,458 24x24), image: IP_Robot.ic_manual_24_80868c
    Rectangle (651,455 339x30), "JOG J4-J6 (MANUAL)"
    RoundedRectangle (615,500 180x64), colour toggle: GVL_Hmi.axJogMinus[4]
    Rectangle (615,500 180x64), "J4 -"
    Rectangle (615,500 180x64)
        tap GVL_Hmi.axJogMinus[4]
    RoundedRectangle (810,500 180x64), colour toggle: GVL_Hmi.axJogPlus[4]
    Rectangle (810,500 180x64), "J4 +"
    Rectangle (810,500 180x64)
        tap GVL_Hmi.axJogPlus[4]
    RoundedRectangle (615,579 180x64), colour toggle: GVL_Hmi.axJogMinus[5]
    Rectangle (615,579 180x64), "J5 -"
    Rectangle (615,579 180x64)
        tap GVL_Hmi.axJogMinus[5]
    RoundedRectangle (810,579 180x64), colour toggle: GVL_Hmi.axJogPlus[5]
    Rectangle (810,579 180x64), "J5 +"
    Rectangle (810,579 180x64)
        tap GVL_Hmi.axJogPlus[5]
    RoundedRectangle (615,658 180x64), colour toggle: GVL_Hmi.axJogMinus[6]
    Rectangle (615,658 180x64), "J6 -"
    Rectangle (615,658 180x64)
        tap GVL_Hmi.axJogMinus[6]
    RoundedRectangle (810,658 180x64), colour toggle: GVL_Hmi.axJogPlus[6]
    Rectangle (810,658 180x64), "J6 +"
    Rectangle (810,658 180x64)
        tap GVL_Hmi.axJogPlus[6]
    RoundedRectangle (1032,434 423x308)
    Image (1056,458 24x24), image: IP_Robot.ic_info_24_80868c
    Rectangle (1092,455 339x30), "ROBOT"
    Ellipse (1056,506 18x18), colour toggle: GVL_HmiView.xJogPermitted
    Rectangle (1089,500 342x29), "Jog permitted", invisible if: NOT (GVL_HmiView.xJogPermitted)
    Rectangle (1089,500 342x29), "Jog locked", invisible if: GVL_HmiView.xJogPermitted
    Ellipse (1056,549 18x18), colour toggle: GVL_HmiView.xRobotMoving
    Rectangle (1089,544 342x29), "Robot moving", invisible if: NOT (GVL_HmiView.xRobotMoving)
    Rectangle (1089,544 342x29), "Robot at rest", invisible if: GVL_HmiView.xRobotMoving
    Ellipse (1056,593 18x18), colour toggle: GVL_Bridge.xVacuumOn
    Rectangle (1089,587 342x29), "Vacuum on", invisible if: NOT (GVL_Bridge.xVacuumOn)
    Rectangle (1089,587 342x29), "Vacuum off", invisible if: GVL_Bridge.xVacuumOn
    Ellipse (1056,636 18x18), colour toggle: GVL_HmiView.axAlarmActive[6]
    Rectangle (1089,631 342x29), "Following error warning", colour toggle: GVL_HmiView.axAlarmActive[6]
    Ellipse (1056,680 18x18), colour toggle: GVL_HmiView.axAlarmActive[7]
    Rectangle (1089,674 342x29), "Following error fault", colour toggle: GVL_HmiView.axAlarmActive[7]
    RoundedRectangle (1473,434 423x308)
    Image (1497,458 24x24), image: IP_Robot.ic_speed_24_80868c
    Rectangle (1533,455 339x30), "SPEED OVERRIDE"
    Rectangle (1497,546 375x24), "Set"
    RoundedRectangle (1497,579 66x66)
    Rectangle (1497,579 66x66), "−"
    Rectangle (1497,579 66x66)
        OnMouseClick: execute { GVL_Hmi.rOverride := LIMIT(0.1, GVL_Hmi.rOverride - 0.1, 1); }
    RoundedRectangle (1575,579 219x66)
    Rectangle (1634,579 101x66), "%.1f", text variable: PRG_HMI_Robot.rV40
    RoundedRectangle (1806,579 66x66)
    Rectangle (1806,579 66x66), "+"
    Rectangle (1806,579 66x66)
        OnMouseClick: execute { GVL_Hmi.rOverride := LIMIT(0.1, GVL_Hmi.rOverride + 0.1, 1); }
    Rectangle (1497,654 375x21), "0.1 – 1"
    RoundedRectangle (150,761 423x200)
    Image (174,785 24x24), image: IP_Robot.ic_machine_24_80868c
    Rectangle (210,782 339x30), "WORST JOINT"
    Rectangle (174,850 143x66), "%.0f", text variable: PRG_HMI_Robot.rV41
    RoundedRectangle (591,761 423x200)
    Image (615,785 24x24), image: IP_Robot.ic_info_24_80868c
    Rectangle (651,782 339x30), "VISION CLASS (0 BOX, 1 JAR, 2 CAN)"
    Rectangle (615,850 143x66), "%.0f", text variable: PRG_HMI_Robot.rV42
    RoundedRectangle (1032,761 423x200)
    Image (1056,785 24x24), image: IP_Robot.ic_info_24_80868c
    Rectangle (1092,782 339x30), "VISION CONFIDENCE"
    Rectangle (1056,850 200x66), "%.2f", text variable: PRG_HMI_Robot.rV43
    RoundedRectangle (1473,761 423x200)
    Image (1497,785 24x24), image: IP_Robot.ic_info_24_80868c
    Rectangle (1533,782 339x30), "VISION POSITION X"
    Rectangle (1497,850 171x66), "%.1f", text variable: PRG_HMI_Robot.rV44
    Rectangle (1677,874 135x37), "mm"
END_VISUALIZATION

// Device/Application/Visu_Alarms
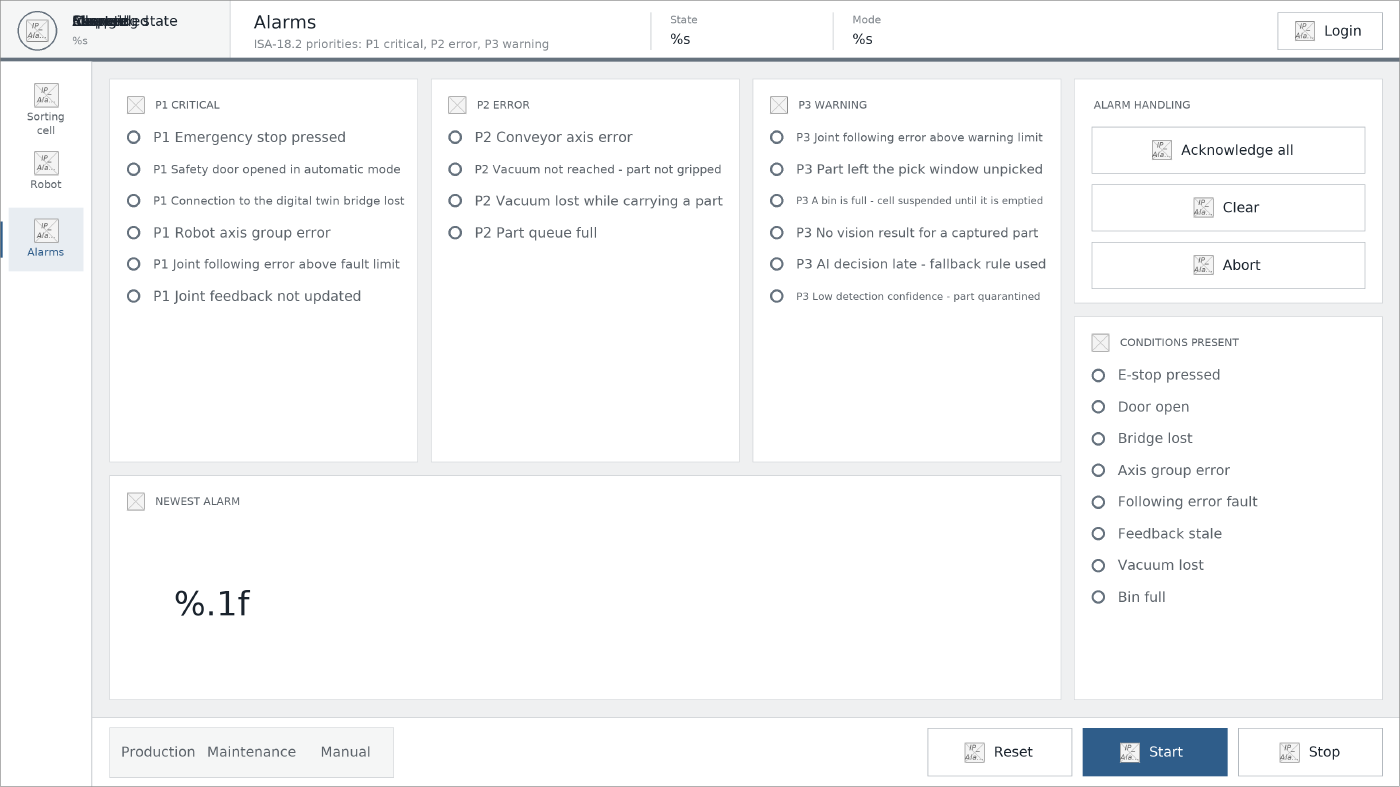
VISUALIZATION Visu_Alarms  // 1920x1080
    Rectangle (0,0 1920x84)
    Rectangle (0,83 1920x1)
    Rectangle (0,0 315x83)
    Rectangle (315,0 1x83)
    Rectangle (0,79 1920x5), invisible if: PRG_HMI_Alarms.iMachine <> 0
    Ellipse (24,15 54x54), invisible if: PRG_HMI_Alarms.iMachine <> 0
    Image (36,27 30x30), invisible if: PRG_HMI_Alarms.iMachine <> 0, image: IP_Alarms.ic_stop_30_66727e
    Rectangle (96,14 198x30), "Stopped", invisible if: PRG_HMI_Alarms.iMachine <> 0
    Rectangle (0,79 1920x5), invisible if: PRG_HMI_Alarms.iMachine <> 1
    Ellipse (24,15 54x54), invisible if: PRG_HMI_Alarms.iMachine <> 1
    Image (36,27 30x30), invisible if: PRG_HMI_Alarms.iMachine <> 1, image: IP_Alarms.ic_fault_30_d72332
    Rectangle (96,14 198x30), "Aborted", invisible if: PRG_HMI_Alarms.iMachine <> 1
    Rectangle (0,79 1920x5), invisible if: PRG_HMI_Alarms.iMachine <> 2
    Ellipse (24,15 54x54), invisible if: PRG_HMI_Alarms.iMachine <> 2
    Image (36,27 30x30), invisible if: PRG_HMI_Alarms.iMachine <> 2, image: IP_Alarms.ic_pause_30_ffbb00
    Rectangle (96,14 198x30), "Suspended", invisible if: PRG_HMI_Alarms.iMachine <> 2
    Rectangle (0,79 1920x5), invisible if: PRG_HMI_Alarms.iMachine <> 3
    Ellipse (24,15 54x54), invisible if: PRG_HMI_Alarms.iMachine <> 3
    Image (36,27 30x30), invisible if: PRG_HMI_Alarms.iMachine <> 3, image: IP_Alarms.ic_warning_30_ffbb00
    Rectangle (96,14 198x30), "Changing state", invisible if: PRG_HMI_Alarms.iMachine <> 3
    Rectangle (0,79 1920x5), invisible if: PRG_HMI_Alarms.iMachine <> 4
    Ellipse (24,15 54x54), invisible if: PRG_HMI_Alarms.iMachine <> 4
    Image (36,27 30x30), invisible if: PRG_HMI_Alarms.iMachine <> 4, image: IP_Alarms.ic_manual_30_2f5d8a
    Rectangle (96,14 198x30), "Manual", invisible if: PRG_HMI_Alarms.iMachine <> 4
    Rectangle (0,79 1920x5), invisible if: PRG_HMI_Alarms.iMachine <> 5
    Ellipse (24,15 54x54), invisible if: PRG_HMI_Alarms.iMachine <> 5
    Image (36,27 30x30), invisible if: PRG_HMI_Alarms.iMachine <> 5, image: IP_Alarms.ic_play_30_66727e
    Rectangle (96,14 198x30), "Execute", invisible if: PRG_HMI_Alarms.iMachine <> 5
    Rectangle (0,79 1920x5), invisible if: PRG_HMI_Alarms.iMachine <> 6
    Ellipse (24,15 54x54), invisible if: PRG_HMI_Alarms.iMachine <> 6
    Image (36,27 30x30), invisible if: PRG_HMI_Alarms.iMachine <> 6, image: IP_Alarms.ic_stop_30_66727e
    Rectangle (96,14 198x30), "Idle", invisible if: PRG_HMI_Alarms.iMachine <> 6
    Rectangle (96,44 198x24), "%s", text variable: GVL_HmiView.sPickStep
    Rectangle (345,11 517x39), "Alarms"
    Rectangle (345,47 517x27), "ISA-18.2 priorities: P1 critical, P2 error, P3 warning"
    Rectangle (892,17 1x51)
    Rectangle (916,15 226x24), "State"
    Rectangle (916,39 226x30), "%s", text variable: PRG_HMI_Alarms.sV1
    Rectangle (1142,17 1x51)
    Rectangle (1166,15 226x24), "Mode"
    Rectangle (1166,39 226x30), "%s", text variable: PRG_HMI_Alarms.sV2
    RoundedRectangle (1752,17 144x51)
    Image (1776,29 27x27), image: IP_Alarms.ic_login_27_1a232d
    Rectangle (1813,17 81x51), "Login"
    Rectangle (1752,17 144x51)
        OnMouseClick:  Type=Login, OpenCentered=True
    Rectangle (126,984 1794x96)
    Rectangle (126,984 1794x1)
    RoundedRectangle (150,998 390x69)
    RoundedRectangle (155,1002 124x60), colour toggle: GVL_HmiPanel.iModeSelect = 1
    Rectangle (155,1002 124x60), "Production", colour toggle: GVL_HmiPanel.iModeSelect = 1
    Rectangle (155,1002 124x60)
        OnMouseClick: execute { GVL_HmiPanel.iModeSelect := 1; }
    RoundedRectangle (283,1002 124x60), colour toggle: GVL_HmiPanel.iModeSelect = 2
    Rectangle (283,1002 124x60), "Maintenance", colour toggle: GVL_HmiPanel.iModeSelect = 2
    Rectangle (283,1002 124x60)
        OnMouseClick: execute { GVL_HmiPanel.iModeSelect := 2; }
    RoundedRectangle (412,1002 124x60), colour toggle: GVL_HmiPanel.iModeSelect = 3
    Rectangle (412,1002 124x60), "Manual", colour toggle: GVL_HmiPanel.iModeSelect = 3
    Rectangle (412,1002 124x60)
        OnMouseClick: execute { GVL_HmiPanel.iModeSelect := 3; }
    RoundedRectangle (1272,999 198x66), colour toggle: GVL_HmiPanel.xReset
    Image (1323,1019 27x27), image: IP_Alarms.ic_reset_27_1a232d
    Rectangle (1360,999 81x66), "Reset"
    Rectangle (1272,999 198x66)
        tap GVL_HmiPanel.xReset
    RoundedRectangle (1485,999 198x66), colour toggle: GVL_HmiPanel.xStart
    Image (1536,1019 27x27), image: IP_Alarms.ic_play_27_ffffff
    Rectangle (1573,999 81x66), "Start"
    Rectangle (1485,999 198x66)
        tap GVL_HmiPanel.xStart
    RoundedRectangle (1698,999 198x66), colour toggle: GVL_HmiPanel.xStop
    Image (1755,1019 27x27), image: IP_Alarms.ic_stop_27_1a232d
    Rectangle (1792,999 69x66), "Stop"
    Rectangle (1698,999 198x66)
        tap GVL_HmiPanel.xStop
    Rectangle (0,84 126x996)
    Rectangle (125,84 1x996)
    Image (47,114 33x33), image: IP_Alarms.ic_home_33_5c636a
    Rectangle (15,150 96x20), "Sorting"
    Rectangle (15,169 96x20), "cell"
    Rectangle (12,99 102x87)
        OnMouseClick:  Assign=Visu_Overview, Type=Assignment
    Image (47,207 33x33), image: IP_Alarms.ic_machine_33_5c636a
    Rectangle (15,243 96x20), "Robot"
    Rectangle (12,192 102x87)
        OnMouseClick:  Assign=Visu_Robot, Type=Assignment
    RoundedRectangle (12,285 102x87)
    RoundedRectangle (0,304 3x49)
    Image (47,300 33x33), image: IP_Alarms.ic_alarm_33_2f5d8a
    Rectangle (15,336 96x20), "Alarms"
    RoundedRectangle (150,108 423x526)
    Image (174,132 24x24), image: IP_Alarms.ic_alarm_24_80868c
    Rectangle (210,129 339x30), "P1 CRITICAL"
    Ellipse (174,179 18x18), colour toggle: GVL_HmiView.axAlarm[1]
    Rectangle (207,174 342x29), "P1 Emergency stop pressed", colour toggle: GVL_HmiView.axAlarm[1]
    Ellipse (174,223 18x18), colour toggle: GVL_HmiView.axAlarm[2]
    Rectangle (207,218 342x29), "P1 Safety door opened in automatic mode", colour toggle: GVL_HmiView.axAlarm[2]
    Ellipse (174,266 18x18), colour toggle: GVL_HmiView.axAlarm[3]
    Rectangle (207,261 342x29), "P1 Connection to the digital twin bridge lost", colour toggle: GVL_HmiView.axAlarm[3]
    Ellipse (174,310 18x18), colour toggle: GVL_HmiView.axAlarm[4]
    Rectangle (207,305 342x29), "P1 Robot axis group error", colour toggle: GVL_HmiView.axAlarm[4]
    Ellipse (174,353 18x18), colour toggle: GVL_HmiView.axAlarm[7]
    Rectangle (207,348 342x29), "P1 Joint following error above fault limit", colour toggle: GVL_HmiView.axAlarm[7]
    Ellipse (174,397 18x18), colour toggle: GVL_HmiView.axAlarm[8]
    Rectangle (207,392 342x29), "P1 Joint feedback not updated", colour toggle: GVL_HmiView.axAlarm[8]
    RoundedRectangle (591,108 423x526)
    Image (615,132 24x24), image: IP_Alarms.ic_alarm_24_80868c
    Rectangle (651,129 339x30), "P2 ERROR"
    Ellipse (615,179 18x18), colour toggle: GVL_HmiView.axAlarm[5]
    Rectangle (648,174 342x29), "P2 Conveyor axis error", colour toggle: GVL_HmiView.axAlarm[5]
    Ellipse (615,223 18x18), colour toggle: GVL_HmiView.axAlarm[9]
    Rectangle (648,218 342x29), "P2 Vacuum not reached - part not gripped", colour toggle: GVL_HmiView.axAlarm[9]
    Ellipse (615,266 18x18), colour toggle: GVL_HmiView.axAlarm[10]
    Rectangle (648,261 342x29), "P2 Vacuum lost while carrying a part", colour toggle: GVL_HmiView.axAlarm[10]
    Ellipse (615,310 18x18), colour toggle: GVL_HmiView.axAlarm[16]
    Rectangle (648,305 342x29), "P2 Part queue full", colour toggle: GVL_HmiView.axAlarm[16]
    RoundedRectangle (1032,108 423x526)
    Image (1056,132 24x24), image: IP_Alarms.ic_warning_24_80868c
    Rectangle (1092,129 339x30), "P3 WARNING"
    Ellipse (1056,179 18x18), colour toggle: GVL_HmiView.axAlarm[6]
    Rectangle (1089,174 342x29), "P3 Joint following error above warning limit", colour toggle: GVL_HmiView.axAlarm[6]
    Ellipse (1056,223 18x18), colour toggle: GVL_HmiView.axAlarm[11]
    Rectangle (1089,218 342x29), "P3 Part left the pick window unpicked", colour toggle: GVL_HmiView.axAlarm[11]
    Ellipse (1056,266 18x18), colour toggle: GVL_HmiView.axAlarm[12]
    Rectangle (1089,261 342x29), "P3 A bin is full - cell suspended until it is emptied", colour toggle: GVL_HmiView.axAlarm[12]
    Ellipse (1056,310 18x18), colour toggle: GVL_HmiView.axAlarm[13]
    Rectangle (1089,305 342x29), "P3 No vision result for a captured part", colour toggle: GVL_HmiView.axAlarm[13]
    Ellipse (1056,353 18x18), colour toggle: GVL_HmiView.axAlarm[14]
    Rectangle (1089,348 342x29), "P3 AI decision late - fallback rule used", colour toggle: GVL_HmiView.axAlarm[14]
    Ellipse (1056,397 18x18), colour toggle: GVL_HmiView.axAlarm[15]
    Rectangle (1089,392 342x29), "P3 Low detection confidence - part quarantined", colour toggle: GVL_HmiView.axAlarm[15]
    RoundedRectangle (150,652 1305x308)
    Image (174,676 24x24), image: IP_Alarms.ic_alarm_24_80868c
    Rectangle (210,673 1221x30), "NEWEST ALARM"
    Rectangle (174,795 171x66), "%.1f", text variable: PRG_HMI_Alarms.rV3
    RoundedRectangle (1473,108 423x308)
    Rectangle (1497,129 375x30), "ALARM HANDLING"
    RoundedRectangle (1497,174 375x64), colour toggle: GVL_HmiPanel.xAckAll
    Image (1580,192 27x27), image: IP_Alarms.ic_check_27_1a232d
    Rectangle (1617,174 194x64), "Acknowledge all"
    Rectangle (1497,174 375x64)
        tap GVL_HmiPanel.xAckAll
    RoundedRectangle (1497,253 375x64), colour toggle: GVL_HmiPanel.xClear
    Image (1637,271 27x27), image: IP_Alarms.ic_reset_27_1a232d
    Rectangle (1674,253 81x64), "Clear"
    Rectangle (1497,253 375x64)
        tap GVL_HmiPanel.xClear
    RoundedRectangle (1497,332 375x64), colour toggle: GVL_HmiPanel.xAbort
    Image (1637,350 27x27), image: IP_Alarms.ic_stop_27_1a232d
    Rectangle (1674,332 81x64), "Abort"
    Rectangle (1497,332 375x64)
        tap GVL_HmiPanel.xAbort
    RoundedRectangle (1473,434 423x526)
    Image (1497,458 24x24), image: IP_Alarms.ic_warning_24_80868c
    Rectangle (1533,455 339x30), "CONDITIONS PRESENT"
    Ellipse (1497,506 18x18), colour toggle: GVL_HmiView.axAlarmActive[1]
    Rectangle (1530,500 342x29), "E-stop pressed", colour toggle: GVL_HmiView.axAlarmActive[1]
    Ellipse (1497,549 18x18), colour toggle: GVL_HmiView.axAlarmActive[2]
    Rectangle (1530,544 342x29), "Door open", colour toggle: GVL_HmiView.axAlarmActive[2]
    Ellipse (1497,593 18x18), colour toggle: GVL_HmiView.axAlarmActive[3]
    Rectangle (1530,587 342x29), "Bridge lost", colour toggle: GVL_HmiView.axAlarmActive[3]
    Ellipse (1497,636 18x18), colour toggle: GVL_HmiView.axAlarmActive[4]
    Rectangle (1530,631 342x29), "Axis group error", colour toggle: GVL_HmiView.axAlarmActive[4]
    Ellipse (1497,680 18x18), colour toggle: GVL_HmiView.axAlarmActive[7]
    Rectangle (1530,674 342x29), "Following error fault", colour toggle: GVL_HmiView.axAlarmActive[7]
    Ellipse (1497,723 18x18), colour toggle: GVL_HmiView.axAlarmActive[8]
    Rectangle (1530,718 342x29), "Feedback stale", colour toggle: GVL_HmiView.axAlarmActive[8]
    Ellipse (1497,767 18x18), colour toggle: GVL_HmiView.axAlarmActive[10]
    Rectangle (1530,761 342x29), "Vacuum lost", colour toggle: GVL_HmiView.axAlarmActive[10]
    Ellipse (1497,810 18x18), colour toggle: GVL_HmiView.axAlarmActive[12]
    Rectangle (1530,805 342x29), "Bin full", colour toggle: GVL_HmiView.axAlarmActive[12]
END_VISUALIZATION
